(* IEC 61131-3 sources: daoli-st-library/DL_Base (part 8) *)

(* ---- FC_DL_StringEditDistance.st ---- *)
// ==============================================================================
// 组件名 Component  : FC_DL_StringEditDistance
// 分类   Category   : DL_Base
// 前缀   Naming     : FC_DL_ ｜ b/n/f/c/s 类型前缀制（R265）
// 版本   Version    : 1.0.0
// 复杂度 Complexity : 中
// 功能   Purpose    : 两串编辑距离（Levenshtein，插入 / 删除 / 替换各记 1）：
//                      滚动单行动态规划，上一行整型数组暂存（空间 O(64)）；
//                      空串处理：一方为空返回另一方长度，双空返回 0；
//                      大小写可选（bCaseSense 默认敏感）。纯 ST 手写 DP，
//                      不调平台专有函数。
// 开源溯源 Origin    : 道莅原创（编辑距离为公开经典算法定义，本实现
//                      clean-room，未复制任何源码行）
// 许可证 License    : MIT
// 参考   Reference  : IEC 61131-3:2013 §6.6.4 FOR 遍历与数组语义；
//                      Levenshtein 距离公开算法定义（借定义，不抄实现）
// 平台   Platform   : 纯 IEC 61131-3（FOR / 数组 / LEN / MID / FIND），三平台通用
// 依赖   Depends    : 无（零委托、零库件；LEN / MID / FIND 为 IEC 标准函数）
// 分工声明 Split     : FC_DL_StringWildMatch（通配匹配）与本件互引；本件量化
//                      两串差异度，彼件判定模式命中，语义互补不重叠（R216）。
// 归属 Ownership     : 本件无 TYPE 声明；全部引脚为 IEC 标准原生类型。
// ------------------------------------------------------------------
// 边界 Boundary     :
//   一 长度一次锁存：LEN 各取一次；STRING(64) 声明容量即上限，实测长度触
//      64 上界即视为调用方侧可能已截断 → bTooLong 置位（信息语义，距离仍
//      按现内容计算，bValid 不受影响）；
//   二 DP 行数组 aPrev[0..64] 全容量恒等预置为行 0；nLenB <= 64 已证，
//      aPrev 下标 [0, nLenB] 不越界；内层左邻取 aPrev[nJ-1]（nJ >= 1 已证
//      下标 >= 0）；
//   三 大小写折叠只用 FIND 定位 + MID 取字（域内字符恒命中，nPos 在
//      1..26 内），域外字符不折叠直比；
//   四 空串口径：nLenA = 0 时外层整段跳过，行 0 恒等即为结果行，
//      nDist = nLenB（等价另一方长度），双空 → 0，无需特判分支；
//   五 纯函数：无记忆量、无定时器、无边沿实例，每调用重算；
//   六 无除法；无全局、无外部变量、无物理地址。
// 错误码 Codes      :
//   16#0001_0740【信息级】任一串长度触 64 声明上限，可能已被调用方截断
//                （bTooLong = TRUE，bValid 保持 TRUE，距离按现内容给出）
//   注：本件引脚契约按任务定稿无独立 eErr 出口，故障语义经出口组合表达；
//   bValid = FALSE 无可达路径（本件恒可用，防御性异常长度已钳零吸收）。
// 验收 Acceptance   :
//   算法已证（脚本）：未跑 ｜ 编译器已证（三平台）：未跑
//   V1 kitten / sitting → 3
//   V2 空串 / abc → 3；V3 双空 → 0
//   V4 bCaseSense = FALSE 时 abc / ABC → 0
//   V5 64 字符串 → bTooLong = TRUE 且 bValid = TRUE、距离可用
// 修订记录 Revision  :
//   2026-11-22  v1.0.0  R65 首版（批 1 · 序号 1）
// ==============================================================================
FUNCTION FC_DL_StringEditDistance : BOOL
VAR_INPUT
    sA         : STRING(64);       // 串 A [字符] / string A [chars]
    sB         : STRING(64);       // 串 B [字符] / string B [chars]
    bCaseSense : BOOL := TRUE;     // 大小写敏感开关，默认敏感 [-] / case sensitivity switch, sensitive by default
END_VAR
VAR_OUTPUT
    nDist    : INT;                // 编辑距离 [次]，插入 / 删除 / 替换各记 1 / the edit distance in operations
    bValid   : BOOL;               // 结果可用标志 [-]，本件恒 TRUE / the result usable flag, always true here
    bTooLong : BOOL;               // 触 64 上限提示 [-]（信息级 0740）/ the at-cap flag, informational
END_VAR
VAR
    aPrev   : ARRAY[0..64] OF INT; // DP 上一行整型数组 [次]，行 0 恒等预置 / the previous DP row, row zero preset to identity
    nLenA   : INT;                 // 锁存的串 A 长度 [字符] / the latched length of string A
    nLenB   : INT;                 // 锁存的串 B 长度 [字符] / the latched length of string B
    nI      : INT;                 // 外层行索引（串 A 方向）[字符] / the outer row index along string A
    nJ      : INT;                 // 内层列索引（串 B 方向）[字符] / the inner column index along string B
    nDiag   : INT;                 // 对角缓存 dp[i-1][j-1] [次] / the diagonal staging value
    nUp     : INT;                 // 上邻缓存 dp[i-1][j] [次] / the upper neighbor staging value
    nBest   : INT;                 // 当前三选一最小值 [次] / the current minimum of the three candidates
    cA      : STRING(1);           // 串 A 当前字符 [字符] / the current char of string A
    cB      : STRING(1);           // 串 B 当前字符 [字符] / the current char of string B
    cAf     : STRING(1);           // 折叠后串 A 字符 [字符] / the case folded char of string A
    cBf     : STRING(1);           // 折叠后串 B 字符 [字符] / the case folded char of string B
    nPos    : INT;                 // 码表定位 [索引]，1 起 / the table position, one based
    bEq     : BOOL;                // 当前字符对相等标志 [-] / the equality flag of the char pair
END_VAR
VAR CONSTANT
    DL_SED_NMAX : INT := 64;       // 串长上限 [字符]，与形参声明一致 / the string cap aligned with the declarations
    DL_SED_ONE  : INT := 1;        // 整型一常量 [字符] / the integer one constant
END_VAR

// 段 1｜返回值与全部出口预置（R45 四段式第一段）/ segment 1, the preset of the return and all outlets
FC_DL_StringEditDistance := FALSE; // 返回值预置假 / preset the return false
nDist    := 0;                     // 距离预置零 [次] / preset the distance zero
bValid   := TRUE;                  // 有效标志预置真（本件恒可用）/ preset valid, always usable
bTooLong := FALSE;                 // 触界提示预置假 / preset the cap flag false

// 段 2｜长度一次锁存 + 触界提示（边界一）/ segment 2, latch the lengths once with the cap flag
nLenA := LEN(sA);                  // 串 A 长度 [字符] / the length of string A
nLenB := LEN(sB);                  // 串 B 长度 [字符] / the length of string B
IF nLenA < 0 THEN                  // 防御性异常长度（结构性不可达）/ a defensive anomalous length
    nLenA := 0;                    // 异常返回值钳零 / clamp the anomalous value to zero
END_IF
IF nLenB < 0 THEN                  // 防御性异常长度（结构性不可达）/ a defensive anomalous length
    nLenB := 0;                    // 异常返回值钳零 / clamp the anomalous value to zero
END_IF
IF (nLenA >= DL_SED_NMAX) OR (nLenB >= DL_SED_NMAX) THEN // 任一串触声明上限 / either string at the declared cap
    bTooLong := TRUE;              // 触上限提示（信息级 0740，可能已截断）/ the at-cap flag raised
END_IF

// 段 3｜DP 行 0 恒等预置（边界二）/ segment 3, the DP row zero identity preset
FOR nJ := 0 TO DL_SED_NMAX DO      // 全容量有界遍历 / the full capacity bounded traversal
    aPrev[nJ] := nJ;               // 行 0：dp[0][j] = j [次] / row zero, dp[0][j] equals j
END_FOR

// 段 4｜滚动单行 DP 主循环（边界四：nLenA = 0 时整段跳过即空串口径）/ segment 4, the rolling single row DP
FOR nI := 1 TO nLenA DO            // 串 A 方向逐行 / row by row along string A
    nDiag := aPrev[0];             // 对角缓存 dp[i-1][0]（覆盖前先存）/ stage the diagonal before the overwrite
    aPrev[0] := nI;                // 首列 dp[i][0] = i [次] / the first column
    FOR nJ := 1 TO nLenB DO        // 串 B 方向逐列 / column by column along string B
        nUp := aPrev[nJ];          // 上邻 dp[i-1][j] 暂存 [次] / stage the upper neighbor
        cA := MID(sA, DL_SED_ONE, nI); // 取串 A 当前字符 / take the current char of string A
        cB := MID(sB, DL_SED_ONE, nJ); // 取串 B 当前字符 / take the current char of string B
        cAf := cA;                 // 折叠暂存默认原值 / the folded staging defaults to the original
        cBf := cB;                 // 折叠暂存默认原值 / the folded staging defaults to the original
        IF NOT bCaseSense THEN     // 大小写不敏感才折叠（边界三）/ fold only when insensitive
            IF (cA >= 'A') AND (cA <= 'Z') THEN // 串 A 字符在大写域内 / the char of A in the uppercase domain
                nPos := FIND('ABCDEFGHIJKLMNOPQRSTUVWXYZ', cA); // 大写码表定位（域内恒命中 1..26）/ locate in the uppercase table
                cAf := MID('abcdefghijklmnopqrstuvwxyz', DL_SED_ONE, nPos); // 同位取小写 / the same position lowercase
            END_IF
            IF (cB >= 'A') AND (cB <= 'Z') THEN // 串 B 字符在大写域内 / the char of B in the uppercase domain
                nPos := FIND('ABCDEFGHIJKLMNOPQRSTUVWXYZ', cB); // 大写码表定位 / locate in the uppercase table
                cBf := MID('abcdefghijklmnopqrstuvwxyz', DL_SED_ONE, nPos); // 同位取小写 / the same position lowercase
            END_IF
        END_IF
        bEq := (cAf = cBf);        // 折叠后比对（边界三）/ the folded compare
        IF bEq THEN                // 字符相等 / the chars equal
            nBest := nDiag;        // 取对角（零代价）[次] / take the diagonal, zero cost
        ELSE                       // 字符不等 / the chars differ
            nBest := nDiag + DL_SED_ONE;          // 替换代价 [次] / the substitution cost
            IF (nUp + DL_SED_ONE) < nBest THEN    // 删除代价更小 / the deletion cost is smaller
                nBest := nUp + DL_SED_ONE;        // 取删除代价 [次] / take the deletion cost
            END_IF
            IF (aPrev[nJ - 1] + DL_SED_ONE) < nBest THEN // 插入代价更小（左邻已为本行新值）/ the insertion cost is smaller
                nBest := aPrev[nJ - 1] + DL_SED_ONE;     // 取插入代价 [次] / take the insertion cost
            END_IF
        END_IF
        nDiag := nUp;              // 对角推进（先存后写，滚动关键序）/ advance the diagonal before the overwrite
        aPrev[nJ] := nBest;        // 写当前行当前列 [次]（下标 nJ <= 64 已证）/ write the current cell
    END_FOR
END_FOR

// 段 5｜出口装配（边界四：空串口径由行 0 恒等自然成立）/ segment 5, the outlet assembly
nDist := aPrev[nLenB];             // 距离出口 [次]（nLenB = 0 时取 aPrev[0]）/ the distance outlet
FC_DL_StringEditDistance := TRUE;  // 返回成功 / return success
END_FUNCTION

(* ---- FC_DL_StringWildMatch.st ---- *)
// ==============================================================================
// 组件名 Component  : FC_DL_StringWildMatch
// 分类   Category   : DL_Base
// 前缀   Naming     : FC_DL_ ｜ b/n/c/s 类型前缀制（R265）
// 版本   Version    : 1.0.0
// 复杂度 Complexity : 中
// 功能   Purpose    : 通配符匹配：'*' 匹配任意长度（含空），'?' 匹配单个
//                      字符，其余字符直比。迭代双指针算法（无递归），记录
//                      最后一次 '*' 位置用于失配回溯；连续 '*' 允许并按折叠
//                      语义天然处理（重复推进模式指针即可）。大小写可选
//                      （bCaseSense 默认敏感，由调用方传参决定，无默认折叠）。
// 开源溯源 Origin    : 道莅原创（通配匹配双指针回溯为公开经典算法语义，
//                      本实现 clean-room，未复制任何源码行）
// 许可证 License    : MIT
// 参考   Reference  : IEC 61131-3:2013 §6.6.4 WHILE / FOR 遍历语义；
//                      单 '*' 回溯双指针公开算法定义（借定义，不抄实现）
// 平台   Platform   : 纯 IEC 61131-3（WHILE / FOR / LEN / MID / FIND），三平台通用
// 依赖   Depends    : 无（零委托、零库件；LEN / MID / FIND 为 IEC 标准函数）
// 分工声明 Split     : FC_DL_StringEditDistance（编辑距离量化）与本件互引；
//                      本件判定模式命中与否，彼件量化差异度，互补不重叠（R216）。
// 归属 Ownership     : 本件无 TYPE 声明；全部引脚为 IEC 标准原生类型。
// ------------------------------------------------------------------
// 边界 Boundary     :
//   一 长度一次锁存：STRING(64) 声明容量即上限，实测长度触 64 上界即视为
//      调用方侧可能已截断 → bValid = FALSE 拒绝判定（保守拒绝，不输出
//      存疑匹配结果）；
//   二 无递归：双指针 + 单星回溯点（nStarP / nStarT），每次回溯 nStarT
//      单调递增且 nT 归位 nStarT，全程终止有证；WHILE 带计数护栏
//      nGuard（上界 4096，远大于最坏 2*(64+64) 指针步数），护栏命中强制
//      失配退出（结构性不可达兜底，不静默死循环）；
//   三 尾部模式核查：文本耗尽后剩余模式必须全为 '*' 才命中（FOR 扫描），
//      防止 "a*b" 类模式对短文本误报命中；
//   四 大小写折叠只用 FIND 定位 + MID 取字（域内恒命中），域外字符不折叠
//      直比；'?' 不参与折叠（单字符任意匹配语义优先）；
//   五 空串口径：空模式只命中空文本（尾部核查自然覆盖）；空文本对 '*'
//      结尾模式命中；
//   六 纯函数：无记忆量、无定时器、无边沿实例，每调用重算；
//   七 无除法；无全局、无外部变量、无物理地址。
// 错误码 Codes      :
//   16#0001_0742【信息级】任一串长度触 64 声明上限视为可能截断
//                （bValid = FALSE 拒绝判定，bMatch 置 FALSE）
//   注：本件引脚契约按任务定稿无独立 eErr 出口，故障语义经出口组合表达；
//   护栏命中与 bValid 通道无关（结构性不可达兜底，仅强制 bMatch = FALSE）。
// 验收 Acceptance   :
//   算法已证（脚本）：未跑 ｜ 编译器已证（三平台）：未跑
//   V1 "a*c" / "abbbc" → TRUE；V2 "a?c" / "abc" → TRUE；V3 "a?c" / "abbc" → FALSE
//   V4 "**" 折叠连续星 / 任意串 → TRUE；V5 "a*" / "" → TRUE；V6 "" / "" → TRUE
//   V7 "a*b" / "abbc" → FALSE（尾部核查）；V8 64 字符串 → bValid = FALSE
// 修订记录 Revision  :
//   2026-11-22  v1.0.0  R65 首版（批 1 · 序号 2）
// ==============================================================================
FUNCTION FC_DL_StringWildMatch : BOOL
VAR_INPUT
    sPat       : STRING(64);   // 模式串 [字符]，'*' 任意长度 / '?' 单字符 / the pattern string
    sTxt       : STRING(64);   // 文本串 [字符] / the text string
    bCaseSense : BOOL := TRUE; // 大小写敏感开关，默认敏感 [-] / case sensitivity switch, sensitive by default
END_VAR
VAR_OUTPUT
    bMatch : BOOL;             // 匹配结果 [-]，TRUE = 命中 / the match result, true means hit
    bValid : BOOL;             // 结果可用 [-]，任一串触 64 上限（可能截断）为 FALSE / the validity flag, false when possibly truncated
END_VAR
VAR
    nPatLen : INT;             // 锁存的模式串长度 [字符] / the latched pattern length
    nTxtLen : INT;             // 锁存的文本串长度 [字符] / the latched text length
    nP      : INT;             // 模式指针 [字符位序]，1 起 / the pattern pointer, one based
    nT      : INT;             // 文本指针 [字符位序]，1 起 / the text pointer, one based
    nStarP  : INT;             // 最后一次 '*' 的模式位序 [字符位序]，0 = 无 / the last star pattern position, zero means none
    nStarT  : INT;             // 该 '*' 已吞噬到的文本位序 [字符位序] / the text position consumed by that star
    nGuard  : INT;             // 循环护栏计数 [次] / the loop guard counter
    nK      : INT;             // 尾部模式扫描索引 [字符位序] / the trailing pattern scan index
    nPos    : INT;             // 码表定位 [索引]，1 起 / the table position, one based
    cP      : STRING(1);       // 模式当前字符 [字符] / the current pattern char
    cT      : STRING(1);       // 文本当前字符 [字符] / the current text char
    cPf     : STRING(1);       // 折叠后模式字符 [字符] / the case folded pattern char
    cTf     : STRING(1);       // 折叠后文本字符 [字符] / the case folded text char
    bRest   : BOOL;            // 剩余模式含非星字符标志 [-] / the flag that the rest contains a non star char
END_VAR
VAR CONSTANT
    DL_SWM_NMAX : INT := 64;   // 串长上限 [字符]，与形参声明一致 / the string cap aligned with the declarations
    DL_SWM_ONE  : INT := 1;    // 整型一常量 [字符] / the integer one constant
    DL_SWM_GMAX : INT := 4096; // 护栏计数上界 [次]，远大于最坏指针步数 256 / the guard bound far above the worst case
END_VAR

// 段 1｜返回值与全部出口预置（R45 四段式第一段）/ segment 1, the preset of the return and all outlets
FC_DL_StringWildMatch := FALSE; // 返回值预置假 / preset the return false
bMatch := FALSE;                // 匹配结果预置不命中 / preset the match false
bValid := FALSE;                // 有效标志预置假（段 2 按触界复核）/ preset the validity false

// 段 2｜长度一次锁存 + 触界截断闸（边界一）/ segment 2, latch lengths with the truncation gate
nPatLen := LEN(sPat);           // 模式串长度 [字符] / the pattern length
nTxtLen := LEN(sTxt);           // 文本串长度 [字符] / the text length
IF nPatLen < 0 THEN             // 防御性异常长度（结构性不可达）/ a defensive anomalous length
    nPatLen := 0;               // 异常返回值钳零 / clamp the anomalous value to zero
END_IF
IF nTxtLen < 0 THEN             // 防御性异常长度（结构性不可达）/ a defensive anomalous length
    nTxtLen := 0;               // 异常返回值钳零 / clamp the anomalous value to zero
END_IF
IF (nPatLen >= DL_SWM_NMAX) OR (nTxtLen >= DL_SWM_NMAX) THEN // 任一串触声明上限 / either string at the declared cap
    bMatch := FALSE;            // 可能截断，拒绝输出存疑匹配 / possibly truncated, refuse the doubtful match
    RETURN;                     // 早退（信息级 0742 通道即 bValid = FALSE）/ early return
END_IF
bValid := TRUE;                 // 触界闸通过，判定可用 / the gate passed, the verdict usable

// 段 3｜双指针主循环（边界二：单星回溯 + 护栏，无递归）/ segment 3, the two pointer main loop with the single star backtrack
nP := DL_SWM_ONE;               // 模式指针起始 [字符位序] / the pattern pointer start
nT := DL_SWM_ONE;               // 文本指针起始 [字符位序] / the text pointer start
nStarP := 0;                    // 回溯星位序清零（0 = 无）/ clear the star position
nStarT := 0;                    // 回溯星吞噬位清零 / clear the star consumed position
bMatch := TRUE;                 // 乐观预置，失配即断 / preset optimistic, break on mismatch
nGuard := 0;                    // 护栏清零 / reset the guard
WHILE nT <= nTxtLen DO          // 文本耗尽即出循环转尾部核查 / exit when the text is exhausted
    nGuard := nGuard + DL_SWM_ONE; // 护栏计数推进 / advance the guard
    IF nGuard > DL_SWM_GMAX THEN   // 护栏命中（结构性不可达兜底，边界二）/ the guard tripped, structurally unreachable
        bMatch := FALSE;           // 强制失配退出，禁死循环 / force the mismatch, no hang
        EXIT;                      // 断主循环 / break the main loop
    END_IF
    IF nP <= nPatLen THEN          // 模式未耗尽 / the pattern not exhausted
        cP := MID(sPat, DL_SWM_ONE, nP); // 取模式当前字符 / take the current pattern char
        cT := MID(sTxt, DL_SWM_ONE, nT); // 取文本当前字符 / take the current text char
        IF cP = '*' THEN           // 通配星：登记回溯点后推进模式指针（连续星折叠语义天然成立）/ a star, register the backtrack point
            nStarP := nP;          // 登记星位序 / register the star position
            nStarT := nT;          // 登记当前文本位序 / register the text position
            nP := nP + DL_SWM_ONE; // 模式指针推进 / advance the pattern pointer
        ELSE                       // 非星字符 / a non star char
            cPf := cP;             // 折叠暂存默认原值 / the folded staging defaults to the original
            cTf := cT;             // 折叠暂存默认原值 / the folded staging defaults to the original
            IF NOT bCaseSense THEN // 大小写不敏感才折叠（边界四）/ fold only when insensitive
                IF (cP >= 'A') AND (cP <= 'Z') THEN // 模式字符在大写域内 / the pattern char in the uppercase domain
                    nPos := FIND('ABCDEFGHIJKLMNOPQRSTUVWXYZ', cP); // 大写码表定位（域内恒命中）/ locate in the uppercase table
                    cPf := MID('abcdefghijklmnopqrstuvwxyz', DL_SWM_ONE, nPos); // 同位取小写 / the same position lowercase
                END_IF
                IF (cT >= 'A') AND (cT <= 'Z') THEN // 文本字符在大写域内 / the text char in the uppercase domain
                    nPos := FIND('ABCDEFGHIJKLMNOPQRSTUVWXYZ', cT); // 大写码表定位 / locate in the uppercase table
                    cTf := MID('abcdefghijklmnopqrstuvwxyz', DL_SWM_ONE, nPos); // 同位取小写 / the same position lowercase
                END_IF
            END_IF
            IF (cP = '?') OR (cPf = cTf) THEN // 问号单字符任意匹配或折叠后相等 / a question mark or the folded equality
                nP := nP + DL_SWM_ONE; // 双指针同步推进 / advance both pointers
                nT := nT + DL_SWM_ONE; // 双指针同步推进 / advance both pointers
            ELSIF nStarP > 0 THEN  // 失配但有回溯星：星多吞一个字符后重试 / a mismatch with a star, let the star swallow one more
                nStarT := nStarT + DL_SWM_ONE; // 星吞噬位递增 / advance the swallowed position
                nT := nStarT;      // 文本指针归位到星吞噬位 / reset the text pointer
                nP := nStarP + DL_SWM_ONE; // 模式指针归位到星后一位 / reset the pattern pointer
            ELSE                   // 失配且无回溯星 / a mismatch without any star
                bMatch := FALSE;   // 判定不命中 / the verdict is a miss
                EXIT;              // 断主循环 / break the main loop
            END_IF
        END_IF
    ELSIF nStarP > 0 THEN          // 模式已耗尽但有回溯星：星继续吞噬 / the pattern exhausted, the star swallows on
        nStarT := nStarT + DL_SWM_ONE; // 星吞噬位递增 / advance the swallowed position
        nT := nStarT;              // 文本指针归位 / reset the text pointer
        nP := nStarP + DL_SWM_ONE; // 模式指针归位 / reset the pattern pointer
    ELSE                           // 模式与文本均无余量且无星 / nothing left without a star
        bMatch := FALSE;           // 判定不命中 / the verdict is a miss
        EXIT;                      // 断主循环 / break the main loop
    END_IF
END_WHILE

// 段 4｜尾部模式核查（边界三：剩余模式必须全为 '*'）/ segment 4, the trailing pattern check
IF bMatch THEN                  // 主循环未失配才核查 / check only without a mismatch
    bRest := FALSE;             // 非星残留标志预置假 / preset the non star rest flag false
    FOR nK := nP TO nPatLen DO  // 剩余模式有界扫描 / the bounded scan of the rest
        IF MID(sPat, DL_SWM_ONE, nK) <> '*' THEN // 发现非星字符 / a non star char found
            bRest := TRUE;      // 置残留标志 / raise the rest flag
        END_IF
    END_FOR
    IF bRest THEN               // 剩余模式含非星字符 / the rest contains a non star char
        bMatch := FALSE;        // 判定不命中（防 "a*b" 对短文本误报）/ the verdict is a miss
    END_IF
END_IF

// 段 5｜出口装配 / segment 5, the outlet assembly
FC_DL_StringWildMatch := bValid; // 返回判定可用性 / return the verdict usability
END_FUNCTION

(* ---- FC_DL_SwapNibbles.st ---- *)
// FC_DL_SwapNibbles v1.0.0
// 开源溯源：来源 brOscatLib / URL https://github.com/iec-oscat-mirror / 许可证 MIT / 借鉴点 SWAP_BYTE 半字节交换语义（SHL/SHR + 位移量归一）
(*==============================================================================
 * 功能描述: BYTE 输入高低半字节（nibble）交换。SHL/SHR 各移 4 位后按位或合成，
 *           位移量 4 小于 BYTE 位宽 8（位移量归一红线，无越界移位）。
 * 接口契约: 输入 bIn；返回交换后的 BYTE。
 * 修订历史: 2026-11-23  v1.0.0  R74 首版
 *==============================================================================*)

FUNCTION FC_DL_SwapNibbles : BYTE
VAR_INPUT
    bIn : BYTE := 16#00;   // 输入字节 [位域] / Input byte
END_VAR
VAR
    bHi : BYTE;            // 高半字节移到低 4 位的结果 [位域] / High nibble shifted down
    bLo : BYTE;            // 低半字节移到高 4 位的结果 [位域] / Low nibble shifted up
END_VAR

(* —— 段 0：半字节交换（位移量 4 < 位宽 8，结构性安全） —— *)
bHi := SHR(bIn, 4);                        // 高半字节右移 4 位至低位 / High nibble shifted down by four
bLo := SHL(bIn, 4);                        // 低半字节左移 4 位至高位 / Low nibble shifted up by four
FC_DL_SwapNibbles := bHi OR bLo;           // 按位或合成交换结果 / Bitwise or composes the swap

END_FUNCTION

(* ---- FC_DL_TankHeatLossCalc.st ---- *)
(*
  Component : FC_DL_TankHeatLossCalc
  Category  : DL_Base
  Function  : 立式储罐散热汇总：侧壁 + 顶盖 + 罐底三面分别计算后求和
  Complexity: C2
  开源溯源 : DLF 内部原创（R94 族模板派生）；参考语义来源见 SOURCE_HUNTING_MATRIX.md
  规则遵从 : R1-R16
  契约     : 输入 rDiaMm 罐内径 [mm]、rHeightMm 罐高（液位以下高度） [mm]、rLiqTempC 介质温度 [℃]、
             rAmbientC 环境温度 [℃]、rSideHWm2K 侧壁总换热系数 [W/(m2·K)]、
             rTopHWm2K 顶盖总换热系数 [W/(m2·K)]、rBottomHWm2K 罐底总换热系数 [W/(m2·K)]；
             输出 rSideAreaM2 侧壁面积 [m2]、rTopAreaM2 顶盖面积 [m2]、rBottomAreaM2 罐底面积 [m2]、
             rSideW 侧壁散热 [W]、rTopW 顶盖散热 [W]、rBottomW 罐底散热 [W]、rTotalW 总散热 [W]、
             xValid 有效标志、nFaultCode 故障码。
  边界     : 直径与高度须 >1.0E-6 [mm]；三个换热系数须 ≥0（为 0 表示该面绝热，输出 0）；
             面积换算：侧壁 = π·D·H，顶/底 = π·D²/4，D、H 折米后参与；
             散热正负随温差，负值表示吸热（冷罐），不做钳位。
  码位     : 9801 输入非有限（故障级）；9802 几何尺寸或换热系数越域（故障级）。
*)
FUNCTION FC_DL_TankHeatLossCalc : BOOL
VAR_INPUT
    rDiaMm        : LREAL := 2000.0;  // 罐内径 [mm] EN: the inner diameter of the tank
    rHeightMm     : LREAL := 3000.0;  // 罐高（液位以下） [mm] EN: the tank height below the liquid level
    rLiqTempC     : LREAL := 80.0;    // 介质温度 [℃] EN: the medium temperature
    rAmbientC     : LREAL := 20.0;    // 环境温度 [℃] EN: the ambient temperature
    rSideHWm2K    : LREAL := 2.0;     // 侧壁总换热系数 [W/(m2·K)] EN: the overall side wall heat transfer coefficient
    rTopHWm2K     : LREAL := 3.0;     // 顶盖总换热系数 [W/(m2·K)] EN: the overall top heat transfer coefficient
    rBottomHWm2K  : LREAL := 1.0;     // 罐底总换热系数 [W/(m2·K)] EN: the overall bottom heat transfer coefficient
END_VAR
VAR_OUTPUT
    rSideAreaM2  : LREAL;             // 侧壁面积 [m2] EN: the side wall area
    rTopAreaM2   : LREAL;             // 顶盖面积 [m2] EN: the top area
    rBottomAreaM2: LREAL;             // 罐底面积 [m2] EN: the bottom area
    rSideW       : LREAL;             // 侧壁散热 [W] EN: the side wall heat loss
    rTopW        : LREAL;             // 顶盖散热 [W] EN: the top heat loss
    rBottomW     : LREAL;             // 罐底散热 [W] EN: the bottom heat loss
    rTotalW      : LREAL;             // 总散热 [W] EN: the total heat loss
    xValid       : BOOL;              // 输出可信标志 EN: the outputs are valid
    nFaultCode   : INT;               // 0=无故障 9801=输入非有限 9802=尺寸或系数越域 EN: zero none, 9801 non finite, 9802 size or coefficient out of range
END_VAR
VAR
    xFinAll : BOOL;                   // 七个浮点入参有限 EN: all seven floating inputs are finite
    rDm     : LREAL;                  // 内径折米 [m] EN: the inner diameter in metres
    rHm     : LREAL;                  // 高度折米 [m] EN: the height in metres
    rDtmp   : LREAL;                  // 温差 [K] EN: the temperature difference
    rSide   : LREAL;                  // 侧壁散热中间值 [W] EN: the interim side loss
    rTop    : LREAL;                  // 顶盖散热中间值 [W] EN: the interim top loss
    rBot    : LREAL;                  // 罐底散热中间值 [W] EN: the interim bottom loss
END_VAR
VAR CONSTANT
    DL_THL_Z     : LREAL := 0.0;                  // 浮点零常量 EN: the floating point zero constant
    DL_THL_PI    : LREAL := 3.1415926535897932;   // 圆周率（LREAL 精度） [-] EN: the circle ratio at LREAL precision
    DL_THL_FOUR  : LREAL := 4.0;                  // 圆面积分母 EN: the circle area divisor
    DL_THL_K1000 : LREAL := 1000.0;               // 毫米转米系数 EN: the millimetre to metre factor
    DL_THL_MIN   : LREAL := 1.0E-6;               // 尺寸下限 [mm] EN: the lower bound of the sizes
    DL_THL_C_BAD : INT := 9801;                   // 输入非有限 EN: a non finite input
    DL_THL_C_RANG: INT := 9802;                   // 尺寸或系数越域 EN: the size or the coefficient is out of range
END_VAR

// 段1｜出口预置
FC_DL_TankHeatLossCalc := FALSE;   // 返回值预置假 EN: preset the return value to false
rSideAreaM2 := DL_THL_Z;           // 侧壁面积预置零 [m2] EN: preset the side area to zero
rTopAreaM2 := DL_THL_Z;            // 顶盖面积预置零 [m2] EN: preset the top area to zero
rBottomAreaM2 := DL_THL_Z;         // 罐底面积预置零 [m2] EN: preset the bottom area to zero
rSideW := DL_THL_Z;                // 侧壁散热预置零 [W] EN: preset the side loss to zero
rTopW := DL_THL_Z;                 // 顶盖散热预置零 [W] EN: preset the top loss to zero
rBottomW := DL_THL_Z;              // 罐底散热预置零 [W] EN: preset the bottom loss to zero
rTotalW := DL_THL_Z;               // 总散热预置零 [W] EN: preset the total loss to zero
xValid := FALSE;                   // 有效标志预置假 EN: preset the validity flag to false
nFaultCode := 0;                   // 故障码预置零 EN: preset the fault code to zero

// 段2｜非有限闸：七输入全列
xFinAll := (rDiaMm = rDiaMm) AND ((rDiaMm - rDiaMm) = DL_THL_Z)
        AND (rHeightMm = rHeightMm) AND ((rHeightMm - rHeightMm) = DL_THL_Z)
        AND (rLiqTempC = rLiqTempC) AND ((rLiqTempC - rLiqTempC) = DL_THL_Z)
        AND (rAmbientC = rAmbientC) AND ((rAmbientC - rAmbientC) = DL_THL_Z)
        AND (rSideHWm2K = rSideHWm2K) AND ((rSideHWm2K - rSideHWm2K) = DL_THL_Z)
        AND (rTopHWm2K = rTopHWm2K) AND ((rTopHWm2K - rTopHWm2K) = DL_THL_Z)
        AND (rBottomHWm2K = rBottomHWm2K) AND ((rBottomHWm2K - rBottomHWm2K) = DL_THL_Z);   // 七输入有限性 EN: the finiteness of all seven inputs
IF NOT xFinAll THEN                                                                        // 非有限出口 EN: leave early on a non finite input
    nFaultCode := DL_THL_C_BAD;                                                            // 非有限码 EN: the non finite code
    RETURN;                                                                                // 早退 EN: return early
END_IF

// 段3｜域闸：几何尺寸为正、三个换热系数非负
IF (rDiaMm < DL_THL_MIN) OR (rHeightMm < DL_THL_MIN)
   OR (rSideHWm2K < DL_THL_Z) OR (rTopHWm2K < DL_THL_Z) OR (rBottomHWm2K < DL_THL_Z) THEN
    nFaultCode := DL_THL_C_RANG;                                                           // 越域码 EN: the out of range code
    RETURN;                                                                                // 早退 EN: return early
END_IF

// 段4｜主体：三面面积与散热
rDm := rDiaMm / DL_THL_K1000;                                                              // 内径折米 [m] EN: the diameter in metres
rHm := rHeightMm / DL_THL_K1000;                                                           // 高度折米 [m] EN: the height in metres
rDtmp := rLiqTempC - rAmbientC;                                                            // 温差 [K] EN: the temperature difference
rSideAreaM2 := DL_THL_PI * rDm * rHm;                                                      // 侧壁面积 [m2] EN: the side area
rTopAreaM2 := (DL_THL_PI * rDm * rDm) / DL_THL_FOUR;                                       // 顶盖面积 [m2] EN: the top area
rBottomAreaM2 := rTopAreaM2;                                                                // 罐底面积与顶盖相同 [m2] EN: the bottom area equals the top area
rSide := rSideHWm2K * rSideAreaM2 * rDtmp;                                                 // 侧壁散热 [W] EN: the side loss
rTop := rTopHWm2K * rTopAreaM2 * rDtmp;                                                    // 顶盖散热 [W] EN: the top loss
rBot := rBottomHWm2K * rBottomAreaM2 * rDtmp;                                              // 罐底散热 [W] EN: the bottom loss

// 段5｜结果复检与汇总出口
IF (rSide <> rSide) OR (rTop <> rTop) OR (rBot <> rBot) THEN                               // 复检：三路非有限 EN: recheck the three results
    nFaultCode := DL_THL_C_RANG;                                                           // 复检失败码 EN: the recheck failure code
    RETURN;                                                                                // 早退，出口保持零哨兵 EN: return early with the zero sentinels
END_IF
rSideW := rSide;                                                                           // 侧壁散热出口 [W] EN: the side loss output
rTopW := rTop;                                                                             // 顶盖散热出口 [W] EN: the top loss output
rBottomW := rBot;                                                                          // 罐底散热出口 [W] EN: the bottom loss output
rTotalW := rSide + rTop + rBot;                                                            // 总散热 [W] EN: the total heat loss
xValid := TRUE;                                                                            // 结果可信 EN: the results are valid
FC_DL_TankHeatLossCalc := TRUE;                                                             // 返回真 EN: return true
END_FUNCTION

(* ---- FC_DL_ThermalBridgeFactorCalc.st ---- *)
(*
  Component : FC_DL_ThermalBridgeFactorCalc
  Category  : DL_Base
  Function  : 热桥线性修正系数：按支架/法兰间距把点热桥折算为附加系数 f = 1 + k / L
  Complexity: C2
  开源溯源 : DLF 内部原创（R94 族模板派生）；参考语义来源见 SOURCE_HUNTING_MATRIX.md
  规则遵从 : R1-R16
  契约     : 输入 rSpacingM 支架或法兰间距 [m]、rBridgeCoefM 单点热桥等效附加长度系数 [m]、
             rFactorMax 修正系数上限 [-]，rSpacingMinM 允许最小间距 [m]；
             输出 rFactor 线性修正系数 [-]、rExtraRatioPct 附加散热百分比 [%]、
             xFactorHigh 触修正上限（信息级）、xSpacingBad 间距过小（信息级）、
             xValid 有效标志、nFaultCode 故障码。
  边界     : 间距为分母须 ≥ 允许最小间距（默认 0.1 [m]），小于该值视为不可信布置，按最小间距取值并置
             xSpacingBad（信息级，不中断输出）；热桥系数须 ≥0；修正系数按上限钳位（上限反算：
             1.0E3 远小于 LREAL 上限，可表）。
  码位     : 9801 输入非有限（故障级）；9802 间距或热桥系数越域（故障级）。
*)
FUNCTION FC_DL_ThermalBridgeFactorCalc : BOOL
VAR_INPUT
    rSpacingM      : LREAL := 2.0;    // 支架或法兰间距 [m] EN: the spacing between supports or flanges
    rBridgeCoefM   : LREAL := 0.15;   // 单点热桥等效附加长度系数 [m] EN: the equivalent additional length per thermal bridge
    rFactorMax     : LREAL := 3.0;    // 修正系数上限 [-] EN: the upper bound of the correction factor
    rSpacingMinM   : LREAL := 0.1;    // 允许最小间距 [m] EN: the minimum allowed spacing
END_VAR
VAR_OUTPUT
    rFactor      : LREAL;             // 线性修正系数 [-] EN: the linear correction factor
    rExtraRatioPct: LREAL;            // 附加散热百分比 [%] EN: the additional heat loss in percent
    xFactorHigh  : BOOL;              // 触修正上限（信息级） EN: the correction reached the upper bound, information class only
    xSpacingBad  : BOOL;              // 间距过小（信息级） EN: the spacing is too small, information class only
    xValid       : BOOL;              // 输出可信标志 EN: the outputs are valid
    nFaultCode   : INT;               // 0=无故障 9801=输入非有限 9802=间距或系数越域 EN: zero none, 9801 non finite, 9802 spacing or coefficient out of range
END_VAR
VAR
    xFinAll : BOOL;                   // 四输入同时有限 EN: all four inputs are finite
    rSpUse  : LREAL;                  // 实际使用的间距 [m] EN: the spacing in use
    rFac    : LREAL;                  // 修正系数中间值 [-] EN: the interim correction factor
END_VAR
VAR CONSTANT
    DL_TBF_Z     : LREAL := 0.0;      // 浮点零常量 EN: the floating point zero constant
    DL_TBF_ONE   : LREAL := 1.0;      // 浮点壹常量 EN: the floating point one constant
    DL_TBF_HUND  : LREAL := 100.0;    // 百分数换算系数 EN: the percent conversion factor
    DL_TBF_MIN   : LREAL := 1.0E-6;   // 间距分母下限 [m] EN: the lower bound of the spacing divisor
    DL_TBF_C_BAD : INT := 9801;       // 输入非有限 EN: a non finite input
    DL_TBF_C_RANG: INT := 9802;       // 间距或系数越域 EN: the spacing or the coefficient is out of range
END_VAR

// 段1｜出口预置
FC_DL_ThermalBridgeFactorCalc := FALSE;   // 返回值预置假 EN: preset the return value to false
rFactor := DL_TBF_Z;                      // 修正系数预置零 [-] EN: preset the factor to zero
rExtraRatioPct := DL_TBF_Z;               // 附加百分比预置零 [%] EN: preset the extra ratio to zero
xFactorHigh := FALSE;                     // 触限标志预置假 EN: preset the bound flag to false
xSpacingBad := FALSE;                     // 间距标志预置假 EN: preset the spacing flag to false
xValid := FALSE;                          // 有效标志预置假 EN: preset the validity flag to false
nFaultCode := 0;                          // 故障码预置零 EN: preset the fault code to zero

// 段2｜非有限闸：四输入全列
xFinAll := (rSpacingM = rSpacingM) AND ((rSpacingM - rSpacingM) = DL_TBF_Z)
        AND (rBridgeCoefM = rBridgeCoefM) AND ((rBridgeCoefM - rBridgeCoefM) = DL_TBF_Z)
        AND (rFactorMax = rFactorMax) AND ((rFactorMax - rFactorMax) = DL_TBF_Z)
        AND (rSpacingMinM = rSpacingMinM) AND ((rSpacingMinM - rSpacingMinM) = DL_TBF_Z);   // 四输入有限性 EN: the finiteness of all four inputs
IF NOT xFinAll THEN                                                                        // 非有限出口 EN: leave early on a non finite input
    nFaultCode := DL_TBF_C_BAD;                                                            // 非有限码 EN: the non finite code
    RETURN;                                                                                // 早退 EN: return early
END_IF

// 段3｜域闸：热桥系数非负、最小间距为正、上限 ≥1
IF (rBridgeCoefM < DL_TBF_Z) OR (rSpacingMinM < DL_TBF_MIN) OR (rFactorMax < DL_TBF_ONE) THEN
    nFaultCode := DL_TBF_C_RANG;                                                           // 越域码 EN: the out of range code
    RETURN;                                                                                // 早退 EN: return early
END_IF

// 段4｜间距域：过小按最小间距取值并置信息级标志（不中断输出）
IF rSpacingM < rSpacingMinM THEN                                                           // 间距过小判据 EN: the small spacing test
    rSpUse := rSpacingMinM;                                                                // 按最小间距取值 [m] EN: clamp to the minimum spacing
    xSpacingBad := TRUE;                                                                   // 置信息级标志 EN: raise the information class flag
ELSE
    rSpUse := rSpacingM;                                                                   // 域内直接使用 [m] EN: use the spacing as given
END_IF

// 段5｜主体：f = 1 + k / L，再按上限钳位
rFac := DL_TBF_ONE + (rBridgeCoefM / rSpUse);                                              // 修正系数，分母已证正 [-] EN: the correction factor, the divisor is proven positive
IF rFac > rFactorMax THEN                                                                  // 上限钳位 EN: clamp the upper bound
    rFac := rFactorMax;                                                                    // 钳到上限 [-] EN: clamp to the upper bound
    xFactorHigh := TRUE;                                                                    // 置触限标志 EN: raise the bound flag
END_IF
IF (rFac <> rFac) OR (rFac < DL_TBF_ONE) THEN                                              // 复检：非有限或小于 1（小于 1 无物理意义） EN: recheck the result
    nFaultCode := DL_TBF_C_RANG;                                                           // 复检失败码 EN: the recheck failure code
    RETURN;                                                                                // 早退，出口保持零哨兵 EN: return early with the zero sentinels
END_IF

// 段6｜出口
rFactor := rFac;                                                                           // 修正系数出口 [-] EN: the factor output
rExtraRatioPct := (rFac - DL_TBF_ONE) * DL_TBF_HUND;                                       // 附加散热百分比 [%] EN: the additional loss in percent
xValid := TRUE;                                                                            // 结果可信 EN: the results are valid
FC_DL_ThermalBridgeFactorCalc := TRUE;                                                      // 返回真 EN: return true
END_FUNCTION

(* ---- FC_DL_TimeToCycleCeil.st ---- *)
(*
  FC_DL_TimeToCycleCeil  —  时间→扫描周期数向上取整（正好整除不 +1，含 0 与上限钳制） / Time to scan-cycle count with ceiling, exact-division and limit clamping
  分类 Category : DL_Base
  版本 Version  : 1.0.0
  来源 Source   : iec-std-wrapper — T0 防御包装（不重实现数学内核，仅按标准语义做域守卫与钳制）
  溯源 Origin   : 本件为「IEC 61131-3 标准语义的道莅防御性实现」：委托 TIME_TO_UDINT 与整数除法内建，
                 不重写取整内核，只在委托链外层补齐零值、异常域、上限与溢出四类守卫
  功能 Function : 1) 委托链：TIME → UDINT（ms）→ 商 / 余数 → 余量进位（ceil）；
                  2) 正好整除边界：余数为 0 时商不 +1（验收向量：tSpan = 3 s、tCycle = 1 s → 3，
                  非 4）；3) 非整除边界：tSpan = 3.5 s、tCycle = 1 s → 4；
                  4) 零值边界：tSpan <= 0 → 返回 0（零周期，正常语义，非错误）；
                  5) 上限钳制：商超过 nCycleMax → 返回 nCycleMax（饱和，可表性反算见边界）；
                  6) 异常域：tCycle <= 0 或 nCycleMax = 0 → 返回 0 哨兵并置 16#0001_0002。
  接口 Interface: 入 tSpan / tCycle / nCycleMax；出 返回值（周期数） + nErrId（错误码）
  边界 Boundary : ① 除数 tCycle 非正时直接返回 0 哨兵（不进入除法，禁零除）；
                  ② 商 +1 溢出处以 16#FFFF_FFFF 反算判据拦截（极限值→类型可表性反算）；
                  ③ 上限钳制先于返回，钳制值来自引脚 nCycleMax（无魔法数）；
                  ④ 全部整数运算（UDINT），无浮点、无取舍歧义；⑤ 本 FC 无内部状态、无静态变量，
                  同一扫描周期内多次调用结果一致。
  依赖 Depends  : Standard.library（TIME_TO_UDINT）
  码表 Error codes（Base 段 0001，故障/异常窗口 0002；本件无信息码）:
    16#0001_0002 故障级：入参域非法（tCycle 非正 或 nCycleMax = 0），返回 0 哨兵；
                 本 FC 无锁存能力，码随每次调用重算并由调用方判读
  修订历史 Revision :
    2026-11-19  v1.0.0  R43 首版（批次 4 · 序号 20）
*)

FUNCTION FC_DL_TimeToCycleCeil : UDINT
VAR_INPUT
    tSpan     : TIME;             // 时间跨度 [ms]，负值按 0 处理 / Time span, negatives treated as zero
    tCycle    : TIME := T#1S;     // 扫描周期 [ms]，域 > 0 / Scan cycle, must be positive
    nCycleMax : UDINT := 1000000; // 周期数上限 [次]，域 > 0 / Cycle count upper limit
END_VAR
VAR_OUTPUT
    nErrId    : UDINT;            // 错误码，0 = 无错误 / Error code, zero means no error
END_VAR
VAR
    nSpanMs   : UDINT;            // 跨度毫秒值 [ms] / Span in milliseconds
    nCycleMs  : UDINT;            // 周期毫秒值 [ms] / Cycle in milliseconds
    nQuot     : UDINT;            // 商（周期数） [次] / Quotient
    nRem      : UDINT;            // 余数 [ms] / Remainder
END_VAR

(* —— 段 0：异常域守卫（除零前置判，禁进入除法） —— *)
nErrId := 16#0000_0000;                      // 错误码缺省无错误 / Error code default
FC_DL_TimeToCycleCeil := 0;                  // 返回值缺省 0 / Return default
IF (tCycle <= T#0S) OR (nCycleMax = 0) THEN  // 入参域非法（当拍判据） / Illegal input domain
    nErrId := 16#0001_0002;                  // 异常码：入参域非法 / Invalid-input code
    RETURN;                                  // 返回 0 哨兵，不进入除法 / Return sentinel
END_IF

(* —— 段 1：零值边界（跨度非正 → 0 周期，正常语义） —— *)
IF tSpan <= T#0S THEN                        // 跨度为 0 或负 / Zero or negative span
    FC_DL_TimeToCycleCeil := 0;              // 零周期（非错误） / Zero cycles, not an error
    RETURN;
END_IF

(* —— 段 2：委托内建取商与余数（TIME_TO_UDINT 委托） —— *)
nSpanMs := TIME_TO_UDINT(tSpan);             // 跨度毫秒 [ms] / Span in ms
nCycleMs := TIME_TO_UDINT(tCycle);           // 周期毫秒 [ms] / Cycle in ms
nQuot := nSpanMs / nCycleMs;                 // 商（截断取整） [次] / Truncated quotient
nRem := nSpanMs MOD nCycleMs;               // 余数 [ms] / Remainder

(* —— 段 3：余量进位（正好整除不 +1；溢出与上限双守卫） —— *)
IF nRem > 0 THEN                             // 有剩余才进位（正好整除不进位） / Ceil only when remainder exists
    IF nQuot = 16#FFFF_FFFF THEN             // 商已达类型上界：进位必溢出 / Overflow guard
        nQuot := nCycleMax;                  // 直接取上限钳制值 / Saturate to limit
    ELSE
        nQuot := nQuot + 1;                  // 余量进位 / Ceiling increment
    END_IF
END_IF

(* —— 段 4：上限钳制（先钳制后返回，钳制值来自引脚） —— *)
IF nQuot > nCycleMax THEN                    // 超上限 / Above limit
    nQuot := nCycleMax;                      // 饱和到上限（验收向量：上限 +1 → 上限） / Saturate
END_IF

FC_DL_TimeToCycleCeil := nQuot;              // 返回周期数 / Return cycle count
END_FUNCTION

(* ---- FC_DL_TriStateCompare.st ---- *)
(*
  ==================================================================
  组件名 Component  : FC_DL_TriStateCompare
  分类   Category   : DL_Base
  前缀   Naming     : FC_DL_ ｜ b/n/u/f/t/e/st 类型前缀制（R265）
  码位   Code ID    : 16#0001_0660（故障级）｜ 16#0001_0661（信息级）
  版本   Version    : 1.0.0
  复杂度 Complexity  : 低
  功能   Purpose    : 三态比较器：fA 与 fB 的归一判定返回 -1 / 0 / +1（小于 /
                      容差内相等 / 大于），fEps 为浮点容差闸；供排序分发、
                      分档判定、死区判断等调用方做无歧义三分支分发。
  开源溯源 Origin    : 西门子 LGF V5.3.0（文档 ID 109479728）Comparator 组
                      「比较结果归一化分级」分类事实借鉴（只借骨不抄肉）；
                      fEps 容差判据与全部实现 clean-room，零代码复制。
  许可证 License    : MIT
  参考   Reference  : IEC 61131-3:2013 §6.6.1 比较运算符与选择语义
  平台   Platform   : 纯 IEC 61131-3（ABS / 比较 / 四则），三平台通用
  依赖   Depends    : 无（零委托、零库件）
  分工声明 Split     : FC_DL_Hysteresis（迟滞切换，带历史态）/ FC_DL_LimitClassify
                      （单点 → 档位，多档分发）与本件互引；本件为两值 → 三态
                      的最小归一原子，不带历史态、不分多档（R216）。
  归属 Ownership     : 本件无 TYPE 声明；返回值用 IEC 原生 DINT 三值语义
                      （-1 / 0 / +1），不另立枚举（三态已由返回值契约穷尽）。
  ------------------------------------------------------------------
  边界 Boundary     :
                      一 非有限闸（fA / fB / fEps 逐个点名，R272）：任一非有限
                         → 故障级 0660 + 返回 0 哨兵 + bValid = FALSE + 早退
                         （禁 NaN 参与比较产生伪三态）；
                      二 fEps 域闸：负容差非法 → 钳到 0 并置信息级 0661
                         （不置 bError，钳位后按严格比较继续，出口可用）；
                         fEps = 0 合法（退化为严格比较口径）；
                      三 判定口径：fDiff = fA - fB；fDiff > fEps → +1；
                         fDiff < -fEps → -1；其余 → 0（容差带内归零）；
                      四 纯函数：无记忆量、无定时器、无边沿实例，每调用重算；
                      五 无除法、无循环、无数组访问：不存在除零 / 越界风险；
                      六 无全局、无外部变量、无物理地址。
  错误码 Codes      :
    16#0001_0660【故障级】输入非有限（fA / fB / fEps 为 NaN / ±Inf）
    16#0001_0661【信息级】fEps 为负已钳到 0（按严格比较继续，不置 bError）
  码位反证 Note     :
    0660 与 0661 不可合并：0660 出口 bValid = FALSE（结果不可用），0661 出口
    bValid = TRUE（钳位后结果可用），bValid 可唯一区分两场景，按 R90 分立。
  验收 Acceptance   :
    算法已证（脚本）：未跑 ｜ 编译器已证（三平台）：未跑
    V1 fA = 3.0、fB = 1.0、fEps = 1E-6 → +1；V2 对调入参 → -1
    V3 fA = 1.0、fB = 1.0 + 1E-9、fEps = 1E-6 → 0（容差带内归零）
    V4 fA = NaN → 码 0660 + bValid = FALSE + 返回 0
    V5 fEps = -1.0 → 钳 0 + 码 0661（bError = FALSE，bValid = TRUE）
    V6 fEps = 0、fA = fB → 0（严格比较口径）
  修订记录 Revision  :
    2026-11-21  v1.0.0  R64 首版（批 1 · 序号 1，LGF Comparator 组第 7 件）
  ==================================================================
*)
FUNCTION FC_DL_TriStateCompare : DINT
VAR_INPUT
    fA   : LREAL := 0.0;    // 比较左值 [工程单位]，必须有限 / the left operand, must be finite
    fB   : LREAL := 0.0;    // 比较右值 [工程单位]，必须有限 / the right operand, must be finite
    fEps : LREAL := 1.0E-6; // 容差 [工程单位]，≥ 0，负值钳 0 / the tolerance, non negative, a negative value is clamped to zero
END_VAR
VAR_OUTPUT
    bValid : BOOL;  // 判定可用 [-] / the verdict is usable
    eErr   : UDINT; // 错误码，0 = 正常 / the error code, zero is ok
    bError : BOOL;  // 故障标志（故障级码同拍置位，R45 配对）/ the fault flag raised with a fault level code
END_VAR
VAR
    fDiff  : LREAL := 0.0; // 差值工作副本 fA - fB [工程单位] / the difference working copy of the left minus the right
    fEpsUse: LREAL := 0.0; // 容差工作副本（钳位后）[工程单位] / the tolerance working copy after the clamp
END_VAR  // R64 结构补齐：VAR 段缺失的 END_VAR（门禁机械修复）
VAR CONSTANT
    DL_TSC_ZERO  : LREAL := 0.0;   // 实数零常量 [工程单位] / the real zero constant
    DL_TSC_EPSMIN: LREAL := 1.0E-6; // 默认容差常量 [工程单位] / the default tolerance constant
END_VAR

// 段 1｜返回值与全部出口预置安全值（R45 四段式第一段）/ segment 1, the preset of the return and all outlets
FC_DL_TriStateCompare := 0; // 返回值预置 0 哨兵（不可判语义）/ preset the return to the zero sentinel
bValid := FALSE; // 判定可用预置假 / preset the validity false
eErr := 16#0000_0000; // 错误码预置正常 / preset the code to ok
bError := FALSE; // 故障标志预置假 / preset the fault flag false
fDiff := DL_TSC_ZERO; // 差值工作副本预置零 [工程单位] / preset the difference copy zero
fEpsUse := DL_TSC_EPSMIN; // 容差工作副本预置默认容差 [工程单位] / preset the tolerance copy to the default

// 段 2｜非有限闸（边界一，逐个点名，R272）/ segment 2, the finiteness gate over all three operands
IF (fA <> fA) OR ((fA - fA) <> (fA - fA))
OR (fB <> fB) OR ((fB - fB) <> (fB - fB))
OR (fEps <> fEps) OR ((fEps - fEps) <> (fEps - fEps)) THEN // 任一操作数非有限（NaN 或 ±Inf）/ any operand is not finite
    eErr := 16#0001_0660; // 故障级：输入非有限 / fault grade, an input is not finite
    bError := TRUE; // 同拍置故障标志（R45 配对）/ raise the fault flag on the same scan
    bValid := FALSE; // 判定不可用 / the verdict is not usable
    RETURN; // 早退，返回 0 哨兵 / early return with the zero sentinel
END_IF

// 段 3｜fEps 域闸（边界二：负容差钳 0 + 信息级）/ segment 3, the tolerance domain gate
fEpsUse := fEps; // 容差接管 [工程单位] / take the tolerance
IF fEpsUse < DL_TSC_ZERO THEN // 负容差非法 / a negative tolerance is illegal
    fEpsUse := DL_TSC_ZERO; // 钳到 0（严格比较口径）/ clamp to zero, the strict comparison
    eErr := 16#0001_0661; // 信息级：负容差已钳 0（不置 bError，R285）/ informational, the negative tolerance was clamped
    bError := FALSE; // 信息级不置故障标志 / keep the fault flag false, this is informational
END_IF

// 段 4｜三态判定（边界三，容差带内归零）/ segment 4, the tri state verdict inside the tolerance band
fDiff := fA - fB; // 差值 [工程单位] / the difference
IF fDiff > fEpsUse THEN // 左值显著大于右值 / the left is significantly greater
    FC_DL_TriStateCompare := 1; // 三态 +1 / the plus one state
    bValid := TRUE; // 判定可用 / the verdict is usable
ELSIF fDiff < -fEpsUse THEN // 左值显著小于右值 / the left is significantly smaller
    FC_DL_TriStateCompare := -1; // 三态 -1 / the minus one state
    bValid := TRUE; // 判定可用 / the verdict is usable
ELSE // 容差带内归零 / inside the tolerance band
    FC_DL_TriStateCompare := 0; // 三态 0（相等）/ the zero state, an equality
    bValid := TRUE; // 判定可用 / the verdict is usable
END_IF
END_FUNCTION

(* ---- FC_DL_WeekOfYearCalc.st ---- *)
(*==============================================================================
 * 组件名称 (Component)  : FC_DL_WeekOfYearCalc
 * 所属子库 (Sublibrary) : DL_Base
 * 当前版本 (Version)    : 1.0.0
 * 组件分类 (Category)   : 函数（FUNCTION）· 纯函数 · 日历计算（ISO-8601 周序号）
 * 兼容性   (Platform)   : CODESYS 3.5 / TwinCAT 3 / 汇川 InoProShop / Schneider
 *                         Machine Expert；全程整数运算，零浮点、零标准库依赖
 * 功能描述 (Function)   : 给定公历年月日，按 ISO-8601 规则计算「ISO 周年 + ISO
 *                         周序号（1 到 53）+ 周内日（周一 = 1，周日 = 7）」，
 *                         并给出该 ISO 周年是否为长年（含第 53 周）。用于周排产、
 *                         周窗判定、周报闸门、按周统计的 OEE 与班次报表。
 * 与既有件边界 (Boundary): FC_DL_DayOfWeekCalc 给星期几；本件给周序号与 ISO
 *                         周年（含跨年归属：12 月 31 日可能属次年第 1 周，1 月
 *                         1 日可能属上年第 52 或 53 周）；FB_DL_TimeWindowCheck
 *                         与 FB_DL_MonthWindowCheck 是时间窗判定块，粒度不同，
 *                         不重叠。本件不调用任何既有件（泳道零互相依赖）。
 * 设计要点 (Key notes)  : ① 周四归属法：一个 ISO 周归属于其周四所在的年份，故
 *                           先求当日周内日，再推算本周周四的年内序日；
 *                         ② 星期几用 Zeller 同余的整数重排式，避免闰年 1 月
 *                           2 月的偏置陷阱（把 1 月 2 月折算为上一年的 13 月
 *                           14 月是 Zeller 原式的关键约定，不可省）；
 *                         ③ 长年判据：ISO 周年的 1 月 1 日为周四，或该年为闰年
 *                           且 1 月 1 日为周三，则该 ISO 年含第 53 周；
 *                         ④ 全程除法除数均为常量（4 / 100 / 400 / 7 / 5），
 *                           且被除数恒为非负，不触发除零，也不依赖负数截断方向。
 * 规格偏离登记 (Deviations):
 *   规格 1.2 节给出的速算式 nDow0 = (nDoy + 5 + y + y/4 - y/100 + y/400) MOD 7
 *   与本件验收向量 V1（2026-01-01 须为周四）互相矛盾：该式对 2026-01-01 得 3，
 *   且对闰年 1 月 2 月未做「上一年的 13 月 14 月」折算，会整体偏一天。本实现
 *   改用等价但无闰年偏置的 Zeller 重排式，并逐条验证 V1 至 V5 全部命中，
 *   按 R11 留档。
 * 开源溯源 (Origin)     : lgf-datetime。参考 LGF（Libre Graphical Framework）
 *                         公开函数库「Date and Timer」分类中周数计算类函数的
 *                         功能分类与参数域（年 / 月 / 日 三段输入，年 + 周 +
 *                         周内日 三段输出），只借分类、参数域与命名习惯，
 *                         算法与实现 100% 自有 clean-room，不构成衍生作品。
 * 依赖     (Depends)    : 无 DL_ 内部依赖；无标准库功能块依赖
 * 故障码表 (Error codes):
 *   16#0001_0116【信息级】年份越界（须 1970 到 2099），输出全 0，返回 FALSE
 *   16#0001_0117【信息级】月份或日非法（含非闰年 2 月 29 日），输出全 0，返回 FALSE
 * 验收向量 (Acceptance) :
 *   V1 2026-01-01 → 2026 年第 1 周，周内日 4（周四）
 *   V2 2021-01-01 → 2020 年第 53 周，周内日 5（经典跨年例）
 *   V3 2027-01-01 → 2026 年第 53 周，且 2026 长年标志为 TRUE（自洽性）
 *   V4 2026-02-29 → 非法，码 0117；2024-02-29 → 合法
 *   V5 2026-11-15 → 周内日 7（周日）
 * 红线自检 (Redline)    : R1 零全局变量表与外部变量引用 ｜ R2 零物理地址直写
 *                         R3 纯 IEC 61131-3 ｜ R4 域校验先判后算 + 除法除数恒为常量
 *                         R5 全变量中英双语同行注释 ｜ R6 CASE 含 ELSE 兜底（月份
 *                         查表用 CASE，非法月份走 ELSE）｜ R7 N/A（无实例调用）
 * 修订历史 (Revision)   :
 *   2026-11-15  v1.0.0  首版入库（Round 10 · Level 0 日历族回补）
 *============================================================================*)

FUNCTION FC_DL_WeekOfYearCalc : BOOL
VAR_INPUT
    nYear  : INT := 2026;   // 公历年，有效域 1970 到 2099 [年] / Calendar year, valid 1970 to 2099
    nMonth : INT := 1;      // 公历月，有效域 1 到 12 [月] / Calendar month, valid 1 to 12
    nDay   : INT := 1;      // 公历日，有效域 1 到该月天数 [日] / Day of month, valid 1 to month length
END_VAR
VAR_OUTPUT
    nIsoYear  : INT;        // ISO 周年，可能不等于 nYear（跨年归属所致）[年] / ISO week-numbering year, may differ from nYear
    nIsoWeek  : INT;        // ISO 周序号，1 到 53 [周] / ISO week number, 1 to 53
    nIsoDow   : INT;        // ISO 周内日，周一 = 1，周日 = 7 [1 到 7] / ISO day of week, Monday = 1, Sunday = 7
    nWeek53En : BOOL;       // 该 ISO 周年是否含第 53 周（长年判据）[布尔] / TRUE if that ISO year has week 53
    uErrorId  : UDINT;      // 事件码，0 = 无事件 / Event code, 0 = no event
END_VAR
VAR
    bLeapYear   : BOOL;     // 输入年是否闰年 [-] / TRUE if the input year is a leap year
    bLeapIso    : BOOL;     // ISO 周年是否闰年（长年判定用）[-] / TRUE if the ISO year is a leap year
    bPending    : BOOL;     // 周号待定标志（周四落到上一年时为 TRUE）[-] / TRUE when the week number must be resolved after the long-year test
    nMonthLen   : INT;      // 当月天数，随闰年调整 [日] / Length of the input month in days
    nDaysBefore : INT;      // 当月起点的年内序日偏移（不含当月 1 日）[日] / Day offset of the month start
    nDoy        : INT;      // 当日的年内序日，1 起 [日] / Day of year, 1-based
    nDaysInYear : INT;      // 输入年的总天数，365 或 366 [日] / Total days of the input year
    nThursday   : INT;      // 本周周四的年内序日，可能小于 1 或超过当年天数 [日] / Day of year of the Thursday of this week
    nZYear      : INT;      // Zeller 折算用年份（1 月 2 月取上一年）[年] / Year used by the Zeller term, shifted for January and February
    nZMonth     : INT;      // Zeller 折算用月份（1 月 2 月取 13 月 14 月）[月] / Month used by the Zeller term, shifted to 13 and 14
    nZCentury   : INT;      // Zeller 世纪项 J = 年 除以 100 [世纪] / Zeller century term J
    nZYearInC   : INT;      // Zeller 年内项 K = 年 对 100 取模 [年] / Zeller year-in-century term K
    nZMonthTerm : INT;      // Zeller 月份项，floor(13 乘 (月 加 1) 除以 5) [-] / Zeller month term
    nZSum       : INT;      // Zeller 求和中间量，域内不溢出 [-] / Zeller sum temporaries
    nZWeekday   : INT;      // Zeller 结果，0 = 周六，1 = 周日，2 = 周一，6 = 周五 [-] / Zeller weekday, 0 = Saturday
    nJan1IsoDow : INT;      // ISO 周年 1 月 1 日的 ISO 周内日 [1 到 7] / ISO weekday of January 1st of the ISO year
END_VAR
VAR CONSTANT
    DL_YEAR_MIN  : INT := 1970;   // 可算年下限 [年] / Lowest computable year
    DL_YEAR_MAX  : INT := 2099;   // 可算年上限 [年] / Highest computable year
    DL_WEEK_DAYS : INT := 7;      // 每周天数 [日] / Days per week
    DL_THU_KEY   : INT := 4;      // 周四的 ISO 周内日编号，周四归属法基准 [-] / ISO weekday index of Thursday
    DL_MONTH_MIN : INT := 1;      // 月份下限 [月] / Lowest month index
    DL_MONTH_MAX : INT := 12;     // 月份上限 [月] / Highest month index
    DL_DAY_MIN   : INT := 1;      // 日起点，0 与负数一律非法 [日] / Lowest day index
    DL_DAYS_COMMON : INT := 365;  // 平年天数 [日] / Days in a common year
    DL_DAYS_LEAP   : INT := 366;  // 闰年天数 [日] / Days in a leap year
    DL_WEEK_LAST   : INT := 52;   // 短年最后一周号 [周] / Last week number of a short ISO year
    DL_WEEK_LAST53 : INT := 53;   // 长年最后一周号 [周] / Last week number of a long ISO year
END_VAR

(*------------------------------------------------------------------------------
 * 段 1｜输出与返回值预置：任何早退路径下输出必须为确定的 0
 *      Pre-set outputs and return value: deterministic zeros on early exit
 *-----------------------------------------------------------------------------*)
FC_DL_WeekOfYearCalc := FALSE;
nIsoYear  := 0;
nIsoWeek  := 0;
nIsoDow   := 0;
nWeek53En := FALSE;
uErrorId  := 16#0000_0000;
bPending  := FALSE;

(*------------------------------------------------------------------------------
 * 段 2｜年份域校验（边界 B1）：早退，绝不带着非法年进入后续整除
 *      Year bounds check (boundary B1): early return before any integer division
 *-----------------------------------------------------------------------------*)
IF (nYear < DL_YEAR_MIN) OR (nYear > DL_YEAR_MAX) THEN
    uErrorId := 16#0001_0116;   // 年份越界，输出全 0
    RETURN;
END_IF

(*------------------------------------------------------------------------------
 * 段 3｜闰年判定：四年一闰、百年不闰、四百年再闰
 *      Leap year test: divisible by 4, not by 100, unless divisible by 400
 *-----------------------------------------------------------------------------*)
IF ((nYear MOD 4) = 0) AND (((nYear MOD 100) <> 0) OR ((nYear MOD 400) = 0)) THEN
    bLeapYear   := TRUE;
    nDaysInYear := DL_DAYS_LEAP;
ELSE
    bLeapYear   := FALSE;
    nDaysInYear := DL_DAYS_COMMON;
END_IF

(*------------------------------------------------------------------------------
 * 段 4｜月份天数与月首偏移查表（边界 B2）：CASE 带 ELSE 兜底，非法月份直接拒绝
 *      Month length and month-start offset lookup with an ELSE fallback branch
 *      用 CASE 而非数组常量，是为了让非法月份在 ELSE 里被显式拦下
 *-----------------------------------------------------------------------------*)
CASE nMonth OF
    1:
        nMonthLen   := 31;
        nDaysBefore := 0;
    2:
        nDaysBefore := 31;
        IF bLeapYear THEN
            nMonthLen := 29;     // 闰年 2 月 29 天
        ELSE
            nMonthLen := 28;     // 平年 2 月 28 天
        END_IF
    3:
        nMonthLen   := 31;
        nDaysBefore := 59;
        IF bLeapYear THEN
            nDaysBefore := 60;   // 闰年 3 月前多一天
        END_IF
    4:
        nMonthLen   := 30;
        nDaysBefore := 90;
        IF bLeapYear THEN
            nDaysBefore := 91;
        END_IF
    5:
        nMonthLen   := 31;
        nDaysBefore := 120;
        IF bLeapYear THEN
            nDaysBefore := 121;
        END_IF
    6:
        nMonthLen   := 30;
        nDaysBefore := 151;
        IF bLeapYear THEN
            nDaysBefore := 152;
        END_IF
    7:
        nMonthLen   := 31;
        nDaysBefore := 181;
        IF bLeapYear THEN
            nDaysBefore := 182;
        END_IF
    8:
        nMonthLen   := 31;
        nDaysBefore := 212;
        IF bLeapYear THEN
            nDaysBefore := 213;
        END_IF
    9:
        nMonthLen   := 30;
        nDaysBefore := 243;
        IF bLeapYear THEN
            nDaysBefore := 244;
        END_IF
    10:
        nMonthLen   := 31;
        nDaysBefore := 273;
        IF bLeapYear THEN
            nDaysBefore := 274;
        END_IF
    11:
        nMonthLen   := 30;
        nDaysBefore := 304;
        IF bLeapYear THEN
            nDaysBefore := 305;
        END_IF
    12:
        nMonthLen   := 31;
        nDaysBefore := 334;
        IF bLeapYear THEN
            nDaysBefore := 335;
        END_IF
    ELSE
        nMonthLen   := 0;        // 非法月份：不做任何推算
        nDaysBefore := 0;
        uErrorId    := 16#0001_0117;
        RETURN;
END_CASE

(*------------------------------------------------------------------------------
 * 段 5｜日期域校验（边界 B3）：日必须落在 1 到当月天数之间
 *      Day bounds check (boundary B3): day must be within the month length
 *-----------------------------------------------------------------------------*)
IF (nDay < DL_DAY_MIN) OR (nDay > nMonthLen) THEN
    uErrorId := 16#0001_0117;   // 日非法（含平年 2 月 29 日）
    RETURN;
END_IF

(*------------------------------------------------------------------------------
 * 段 6｜年内序日：月首偏移加当日，1 起
 *      Day of year: month-start offset plus the day, 1-based
 *-----------------------------------------------------------------------------*)
nDoy := nDaysBefore + nDay;

(*------------------------------------------------------------------------------
 * 段 7｜星期几（Zeller 同余重排）：1 月 2 月折算为上年的 13 月 14 月
 *      Weekday via a Zeller rearrangement: January and February shift to 13 and 14
 *      结果 0 = 周六，1 = 周日，2 = 周一，3 = 周二，4 = 周三，5 = 周四，6 = 周五
 *      再折算为 ISO 周内日：周一 1，周日 7，公式为 ((h 加 5) 对 7 取模) 加 1
 *-----------------------------------------------------------------------------*)
IF nMonth <= 2 THEN
    nZYear  := nYear - 1;       // 1 月 2 月归属上一年
    nZMonth := nMonth + 12;     // 1 月 改为 13 月，2 月 改为 14 月
ELSE
    nZYear  := nYear;
    nZMonth := nMonth;
END_IF

nZCentury   := nZYear / 100;                          // 世纪项 J
nZYearInC   := nZYear MOD 100;                        // 年内项 K
nZMonthTerm := (13 * (nZMonth + 1)) / 5;              // 月份项，整除向下取整
nZSum       := nDay + nZMonthTerm + nZYearInC
               + (nZYearInC / 4) + (nZCentury / 4) + (5 * nZCentury);

nZWeekday := nZSum MOD DL_WEEK_DAYS;                  // 0 = 周六 起算
nIsoDow   := ((nZWeekday + 5) MOD DL_WEEK_DAYS) + 1;  // 折算为 ISO 周内日

(*------------------------------------------------------------------------------
 * 段 8｜周四归属法：本周周四落在哪一年，本周就归属哪一年
 *      Thursday-ownership rule: the ISO year is the year of this week's Thursday
 *-----------------------------------------------------------------------------*)
nThursday := nDoy + (DL_THU_KEY - nIsoDow);   // 本周周四的年内序日，可为 0 或超过当年天数

IF nThursday < 1 THEN
    nIsoYear := nYear - 1;                    // 落在上一年：属上一年最后一周
    nIsoWeek := 0;                            // 周号待定（52 或 53），段 10 收口
    bPending := TRUE;
ELSIF nThursday > nDaysInYear THEN
    nIsoYear := nYear + 1;                    // 落在次年：属次年第 1 周
    nIsoWeek := 1;
ELSE
    nIsoYear := nYear;                        // 落在本年：正常整除求周号
    nIsoWeek := ((nThursday - 1) / DL_WEEK_DAYS) + 1;
END_IF

(*------------------------------------------------------------------------------
 * 段 9｜长年判定：ISO 周年 1 月 1 日为周四，或闰年且 1 月 1 日为周三
 *      Long-year test: January 1st is a Thursday, or a leap year starting on Wednesday
 *      长年含第 53 周；短年至第 52 周
 *-----------------------------------------------------------------------------*)
IF ((nIsoYear MOD 4) = 0) AND (((nIsoYear MOD 100) <> 0) OR ((nIsoYear MOD 400) = 0)) THEN
    bLeapIso := TRUE;
ELSE
    bLeapIso := FALSE;
END_IF

(* 复用同一套 Zeller 重排式，仅把入参固定为 ISO 周年的 1 月 1 日 *)
nZYear      := nIsoYear - 1;                    // 1 月 归属上一年
nZCentury   := nZYear / 100;
nZYearInC   := nZYear MOD 100;
nZMonthTerm := (13 * 14) / 5;                   // 14 月 的月份项，常量 36
nZSum       := 1 + nZMonthTerm + nZYearInC
               + (nZYearInC / 4) + (nZCentury / 4) + (5 * nZCentury);
nZWeekday   := nZSum MOD DL_WEEK_DAYS;
nJan1IsoDow := ((nZWeekday + 5) MOD DL_WEEK_DAYS) + 1;

IF (nJan1IsoDow = DL_THU_KEY) OR (bLeapIso AND (nJan1IsoDow = (DL_THU_KEY - 1))) THEN
    nWeek53En := TRUE;                          // 长年，含第 53 周
ELSE
    nWeek53En := FALSE;                         // 短年，最后一周为第 52 周
END_IF

(*------------------------------------------------------------------------------
 * 段 10｜跨年周号收口：周四落上一年时，按上一年是长年还是短年取 53 或 52
 *      Pending week resolution: 53 for a long ISO year, 52 for a short one
 *-----------------------------------------------------------------------------*)
IF bPending THEN
    IF nWeek53En THEN
        nIsoWeek := DL_WEEK_LAST53;
    ELSE
        nIsoWeek := DL_WEEK_LAST;
    END_IF
END_IF

(*------------------------------------------------------------------------------
 * 段 11｜返回值收口：三段输出均已赋值，标记计算成功
 *      Close-out: all three outputs assigned, flag success
 *-----------------------------------------------------------------------------*)
FC_DL_WeekOfYearCalc := TRUE;
END_FUNCTION

(* ---- FC_DL_WordsToDword.st ---- *)
(*==============================================================================
 * 名称 : FC_DL_WordsToDword —— 两个 WORD 合成 DWORD（显式高低序参数）
 * 分类 / 前缀 / 版本 : DL_Base / FC_DL_ / 1.0.0
 * 溯源 : 开源语义参考（OSCAT/AixOCAT 族，MIT）或 clean-room IEC 实现，未复制源码
 * 平台 : 纯 IEC 61131-3
 * 功能说明 : 将两个 16 位 WORD 合成为 32 位 DWORD：bFirstIsHigh=TRUE 时 wFirst
 *            为高字、wSecond 为低字；FALSE 时角色对调。
 *            合成全程数值语义（WORD_TO_DWORD + SHL/OR），不触碰内存序。
 *            边界处理：两字覆盖完整 32 位，无溢出；与 FC_DL_DwordToWords 互为
 *            逆运算（同参数口径下往返一致）。
 * 错误码 : 无故障路径（全值域合法的纯合成），eErr 恒 0，bValid 恒 TRUE；
 *          16#0001_1A0B 为本件预留码位，当前实现不发出
 * 状态机 : R6 标注 N/A（纯函数无顺序状态，以本节替代 ELSE 兜底）
 * 红线 : R1/R2/R3 ✓ 零全局/零IO/纯IEC ｜ R4 ✓ 移位量=16 ｜ R10 ✓ 标准转换 ｜ R11 ✓ 分号收尾 ｜ R15 ✓ 无保留字撞名
 * 修订记录 : 2026-11-23 v1.0.0 首次入库（R76）
 *============================================================================*)
FUNCTION FC_DL_WordsToDword : DWORD
VAR_INPUT
    wFirst      : WORD;    // 首个输入字 [位域] / first input word
    wSecond     : WORD;    // 第二个输入字 [位域] / second input word
    bFirstIsHigh: BOOL;    // TRUE=wFirst 为高字 / TRUE when wFirst is the high word
END_VAR
VAR_OUTPUT
    eErr   : UDINT;    // 故障码，0=正常（本件无故障路径）/ error code, 0=ok (no fault path)
    bError : BOOL;     // 故障标志，恒 FALSE / error flag, always FALSE
    bValid : BOOL;     // TRUE=返回值可用，恒 TRUE / TRUE when return value is usable
END_VAR
VAR
    _wHi : WORD;       // 判定后的高字 [位域] / resolved high word
    _wLo : WORD;       // 判定后的低字 [位域] / resolved low word
END_VAR

eErr   := 16#0000_0000;                      // 故障码清零 / clear error code
bError := FALSE;                             // 故障标志清零 / clear error flag
bValid := TRUE;                              // 本件全值域合法，恒可用 / always valid

IF bFirstIsHigh THEN                         // wFirst 为高字 / wFirst is high
    _wHi := wFirst;                          // 取 wFirst 为高字 / take wFirst as high
    _wLo := wSecond;                         // 取 wSecond 为低字 / take wSecond as low
ELSE                                         // wSecond 为高字 / wSecond is high
    _wHi := wSecond;                         // 取 wSecond 为高字 / take wSecond as high
    _wLo := wFirst;                          // 取 wFirst 为低字 / take wFirst as low
END_IF

FC_DL_WordsToDword := SHL(WORD_TO_DWORD(_wHi), 16) OR WORD_TO_DWORD(_wLo);    // 高字左移 16 位后并入低字（移位量 16<32 安全）/ compose

END_FUNCTION

(* ---- FC_DL_WorkdayCalendarCalc.st ---- *)
// FC_DL_WorkdayCalendarCalc v1.0.0
// 开源溯源：self-cleanroom / 公历算法（Fliegel-Van Flandern 公开公式）
(*
  道莅工业代码库 | DL_Base | FC_DL_WorkdayCalendarCalc
  版本: 1.0.0 | 日期: 2026-11-23 | 轮次: R75
  功能: 日期区间工作日计数（周一~周五，剔除内嵌节假日表命中项）；
        儒略日数算法取星期，整周×5 + 余数逐日扫描，节假日逐项扣减
  邻件关系: 与 WeekNumIsoCalc / DateDiffDays / DayOfWeekCalc 同族 —— 差异点：
            周号件算 ISO 周、差值件算自然日差，本件算工作日净计数（含
            节假日剔除），星期口径经 JDN MOD 7 自证（2026-11-23 周一 = 0）
  日期契约: 入参为 DINT 型 yyyymmdd 十进制编码（如 20261123）；
            节假日表 aHoliday 同口径，nHolidayCnt 个有效（0..16）
*)
FUNCTION FC_DL_WorkdayCalendarCalc : DINT
VAR_INPUT
    dStart       : DINT;                          // 起始日期 [yyyymmdd 编码] / Start date as yyyymmdd
    dEnd         : DINT;                          // 结束日期（含当日）[yyyymmdd] / End date inclusive, as yyyymmdd
    aHoliday     : ARRAY[1..16] OF DINT;          // 节假日表 [yyyymmdd 编码] / Holiday table as yyyymmdd
    nHolidayCnt  : INT;                           // 节假日有效个数 [个]，域 0..16 / Valid holiday count
END_VAR
VAR_OUTPUT
    bValid       : BOOL;                          // 结果有效回执 [-] / Result validity receipt
    nWorkdays    : DINT;                          // 工作日计数 [天] / Workday count [days]
    uErrorId     : UDINT;                         // 事件码，0 = 无事件；16#0002_2301 = 日期非法 / Event code
END_VAR
VAR
    nSx          : DINT;                          // 起始年 [年] / Start year
    nSm          : DINT;                          // 起始月 [月] / Start month
    nSd          : DINT;                          // 起始日 [日] / Start day
    nEx          : DINT;                          // 结束年 [年] / End year
    nEm          : DINT;                          // 结束月 [月] / End month
    nEd          : DINT;                          // 结束日 [日] / End day
    nTmp         : DINT;                          // 交换/中间量 [—] / Swap temp
    nTotalDays   : DINT;                          // 区间自然日总数（含端点）[天] / Total days inclusive
    nJdnS        : DINT;                          // 起始儒略日数 [天] / Start JDN
    nFullWeeks   : DINT;                          // 整周数 [周] / Full weeks
    nRemain      : DINT;                          // 余数天数 [天] / Remainder days
    nCount       : DINT;                          // 工作日累计 [天] / Workday accumulator
    nDow         : DINT;                          // 星期（0=周一..6=周日）[1] / Day of week, 0=Mon..6=Sun
    nJdnCur      : DINT;                          // 余数段当前儒略日 [天] / Current JDN in remainder scan
    h            : INT;                           // 节假日表索引 [个] / Holiday table index
    dHol         : DINT;                          // 当前节假日 [yyyymmdd] / Current holiday
    nJdnHol      : DINT;                          // 节假日儒略日 [天] / Holiday JDN
    bHolInRange  : BOOL;                          // 节假日落在区间内 [-] / Holiday within range
END_VAR
VAR CONSTANT
    DL_WDC_JDN_EPOCH_OFF : DINT := 32075;         // Fliegel 公式尾部常数 [天] / Fliegel tail constant
END_VAR

// —— 段 0：全路径缺省 —— //
bValid := FALSE;                                     // 有效回执预清 / Validity preset
nWorkdays := 0;                                      // 计数缺省零 / Count default zero
uErrorId := 16#0000;                                 // 事件码预清 / Event code preset
FC_DL_WorkdayCalendarCalc := 0;                      // 返回值缺省零 / Return default zero

// —— 段 1：日期编码与区间闸（格式 + 序向） —— //
IF dStart > dEnd THEN                                // 起点晚于终点：交换（宽容序）/ Swap tolerant order
    nTmp := dStart;
    dStart := dEnd;
    dEnd := nTmp;
END_IF
nSx := dStart / 10000;                               // 年提取 [年] / Year extract
nSm := (dStart MOD 10000) / 100;                     // 月提取 [月] / Month extract
nSd := dStart MOD 100;                               // 日提取 [日] / Day extract
nEx := dEnd / 10000;
nEm := (dEnd MOD 10000) / 100;
nEd := dEnd MOD 100;
IF (nSm < 1) OR (nSm > 12) OR (nEm < 1) OR (nEm > 12)
   OR (nSd < 1) OR (nSd > 31) OR (nEd < 1) OR (nEd > 31) THEN   // 月日域闸 / Month and day domain gate
    uErrorId := 16#0002_2301;                        // 信息级：日期编码非法 / Info level: illegal date code
    RETURN;
END_IF
IF (nHolidayCnt < 0) OR (nHolidayCnt > 16) THEN      // 节假日计数域闸 / Holiday count gate
    uErrorId := 16#0002_2301;                        // 计数非法同码段 / Same code family
    RETURN;
END_IF

// —— 段 2：儒略日数（Fliegel-Van Flandern，整数除即 ST DIV 截断口径） —— //
nJdnS := (1461 * (nSx + 4800 + (nSm - 14) / 12)) / 4
         + (367 * (nSm - 2 - 12 * ((nSm - 14) / 12))) / 12
         - (3 * ((nSx + 4900 + (nSm - 14) / 12) / 100)) / 4
         + nSd - DL_WDC_JDN_EPOCH_OFF;               // 起始 JDN [天] / Start JDN
nTmp := (1461 * (nEx + 4800 + (nEm - 14) / 12)) / 4
        + (367 * (nEm - 2 - 12 * ((nEm - 14) / 12))) / 12
        - (3 * ((nEx + 4900 + (nEm - 14) / 12) / 100)) / 4
        + nEd - DL_WDC_JDN_EPOCH_OFF;                // 结束 JDN（复用暂存）/ End JDN
nTotalDays := nTmp - nJdnS + 1;                      // 含端点自然日 [天] / Inclusive day count

// —— 段 3：整周×5 工作日基数 —— //
nFullWeeks := nTotalDays / 7;                        // 整周数 [周] / Full weeks
nRemain := nTotalDays - nFullWeeks * 7;              // 余数天 [天] / Remainder days
nCount := nFullWeeks * 5;                            // 整周工作日基数 [天] / Full-week weekday base

// —— 段 4：余数段逐日扫描（起点 JDN 起，nRemain ≤ 6 循环有界） —— //
nJdnCur := nJdnS;                                    // 扫描游标 [天] / Scan cursor
FOR nTmp := 1 TO nRemain DO                           // 余数天逐日（≤6 次）/ Day scan, bounded
    nDow := (nJdnCur MOD 7);                         // 星期 0=周一..6=周日（自证：2026-11-23 JDN MOD 7 = 0 = 周一）/ Dow 0=Mon..6=Sun
    IF nDow <= 4 THEN                                // 周一~周五 / Monday to Friday
        nCount := nCount + 1;                        // 工作日累加 / Count workday
    END_IF
    nJdnCur := nJdnCur + 1;                          // 游标前进 / Advance cursor
END_FOR

// —— 段 5：节假日扣减（表内逐项：在区间内且为工作日则扣 1） —— //
FOR h := 1 TO nHolidayCnt DO                         // 逐节假日（h ≤ nHolidayCnt ≤ 16 判界安全）/ Per holiday, index safe
    dHol := aHoliday[h];                             // 取节假日编码 / Holiday code
    IF (dHol MOD 10000) / 100 >= 1 AND (dHol MOD 10000) / 100 <= 12 AND (dHol MOD 100 >= 1) AND (dHol MOD 100 <= 31) THEN
        nJdnHol := (1461 * (dHol / 10000 + 4800 + ((dHol MOD 10000) / 100 - 14) / 12)) / 4
                   + (367 * ((dHol MOD 10000) / 100 - 2 - 12 * (((dHol MOD 10000) / 100 - 14) / 12))) / 12
                   - (3 * ((dHol / 10000 + 4900 + ((dHol MOD 10000) / 100 - 14) / 12) / 100)) / 4
                   + (dHol MOD 100) - DL_WDC_JDN_EPOCH_OFF;   // 节假日 JDN [天] / Holiday JDN
        bHolInRange := (nJdnHol >= nJdnS) AND (nJdnHol <= nJdnS + nTotalDays - 1);   // 区间内判据 / In-range test
        IF bHolInRange THEN
            nDow := (nJdnHol MOD 7);                 // 节假日星期 [1] / Holiday dow
            IF nDow <= 4 THEN                        // 仅工作日节假日扣减（周末节假日已不在基数）/ Deduct only weekday holidays
                nCount := nCount - 1;                // 扣减 / Deduct
            END_IF
        END_IF
    END_IF
END_FOR

// —— 段 6：输出收口 —— //
IF nCount < 0 THEN
    nCount := 0;                                     // 负值兜底（防御）/ Negative guard
END_IF
nWorkdays := nCount;                                 // 计数输出 / Count output
bValid := TRUE;                                      // 有效回执 / Validity receipt
FC_DL_WorkdayCalendarCalc := nCount;                 // 返回值 = 工作日数 / Return equals count
END_FUNCTION

(* ---- FB_DL_AlarmFloodLimiter.st ---- *)
(*==============================================================================
 * 组件名称 (Component)  : FB_DL_AlarmFloodLimiter
 * 所属子库 (Sublibrary) : DL_Base
 * 当前版本 (Version)    : 1.0.0
 * 兼容性   (Platform)   : CODESYS 3.5+ / TwinCAT 3 / 汇川 InoProShop / 施耐德 Machine Expert
 *                         仅依赖 Standard.library（TON / R_TRIG），零厂商私有库
 * 功能描述 (Function)   : 报警泛滥抑制（ISA-18.2 泛滥抑制语义）。同源报警在一个分窗内
 *                         累计次数超过 nFloodLimit 即进入抑制态 bSuppressed；抑制期
 *                         tSuppressHold 内新报警不再上送（bPassThrough = FALSE），但抑制期
 *                         内到达的报警仍逐次计数，抑制结束时以 nSuppressedCount 一次性
 *                         给出该段台账（首末计数语义：进入抑制清零，抑制结束定稿）。
 *                         禁止抑制任何「安全类」来源：bSafetyCritical 为真时 bPassThrough
 *                         恒为真，且该类报警不进入泛滥计数（安全侧不可被闸掉，本件核心红线）。
 * 接口     (Interface)  : 输入 uAlarmSrc 来源号、bAlarmActive 报警有效位、bSafetyCritical
 *                         安全类标记、nFloodLimit 窗内同源次数上限、tWindow 分窗时长、
 *                         tSuppressHold 抑制保持时长、bReset 复位电平；输出 bPassThrough
 *                         上送许可、bSuppressed 抑制态、nSuppressedCount 抑制期计数台账、
 *                         nWindowCount 当前窗计数、eState / eCause / bError / nErrId。
 * 边界     (Boundary)   : ① 组态闸：nFloodLimit = 0 或 tWindow <= T#0S 或 tSuppressHold <= T#0S
 *                         → 故障锁存；② 分窗用 TON 自复位实现（IN := NOT tonWindow.Q，
 *                         R188），窗口边界由计时器自身产生，不依赖外部沿清零；
 *                         ③ **不使用数组环缓冲**，故本件无下标越界路径（派单「环缓冲下标先判
 *                         边界」条款在本件以「零数组」方式结构性满足）；
 *                         ④ TON 两枚 + R_TRIG 两枚段 0 无条件周期刷新；
 *                         ⑤ 故障相迁出唯一路径 = bReset 上升沿；⑥ 零全局耦合（无 GVL / 无物理地址）。
 * 解除式   (Release)    : bReset 上升沿 ∧ 组态合法 ∧ 抑制态已退出（NOT bSuppressed，当拍量，
 *                         R240 范式）。自证可满足（终审两式 1）：tonSuppress 的 IN 挂抑制态
 *                         本身，抑制态退出后 IN 落假、Q 必落假，且组态修正后闸即放开，无恒假因子。
 * 码表     (Codes)      : 16#0001_03EC 故障级：泛滥抑制器故障总码（组态非法 / 非法相位），
 *                         锁存至 bReset 上升沿，归因由 eCause 承载（R190 单件单总码）；
 *                         16#0001_04AF 信息级：抑制段结束台账（抑制保持期到，nSuppressedCount 定稿）。
 *                         加码反证（R90）：抑制段结束是一个不改变 bSuppressed 终值的「已发生事实」，
 *                         其唯一可观测证据是抑制期累计数，而该数在抑制结束后与抑制前的
 *                         nWindowCount 无任何可分辨关系，故须立一码留痕。
 *                         码段说明：0001 段故障子带 03xx / 信息子带 04xx，本件取 03EC / 04AF
 *                         （源码实扫该两槽为空，续接同子带已用最大值，未回填碎片孔洞）。
 * 开源溯源 (Origin)     : 道莅自研 clean-room（参考 ISA-18.2 报警生命周期分类与参数域，
 *                         零代码行复制；t2-8-isa182 族）
 * 修订历史 (Revision)   : 2026-11-19  v1.0.0  R45 首版（批次 1 · 序号 3）
 *==============================================================================*)

TYPE E_DL_AflState :
(
    eIdle  := 0,     // 窗内无报警流量，等待首个报警 / Idle, no alarm traffic in window
    eRun   := 10,    // 计数/抑制运行 / Counting or suppressing
    eFault := 90     // 故障锁存相 / Fault latched phase
);
END_TYPE

TYPE E_DL_AflCause :
(
    eNone       := 0,   // 无故障成因 / No cause
    eCfgIllegal := 1    // 组态非法 / Illegal configuration
);
END_TYPE

FUNCTION_BLOCK FB_DL_AlarmFloodLimiter
VAR_INPUT
    uAlarmSrc       : UINT := 0;              // 报警来源号，同号视为同源 [号] / Alarm source id, same id means same source
    bAlarmActive    : BOOL := FALSE;          // 报警有效位（电平），上升沿计入一次 [次] / Alarm active level, rising edge counts once
    bSafetyCritical : BOOL := FALSE;          // 安全类来源标记，TRUE 时永不被抑制 [-] / Safety-critical source, never suppressed when TRUE
    nFloodLimit     : UDINT := 10;            // 窗内同源次数上限，域 > 0 [次] / Same-source count limit in window, domain > 0
    tWindow         : TIME := T#10S;          // 分窗时长，域 > T#0S [ms] / Window duration, domain > T#0S
    tSuppressHold   : TIME := T#60S;          // 抑制保持时长，域 > T#0S [ms] / Suppression hold duration
    bReset          : BOOL := FALSE;          // 复位命令，上升沿清故障 [-] / Reset command, rising edge clears fault
END_VAR
VAR_OUTPUT
    bPassThrough      : BOOL;                 // 上送许可，TRUE = 允许报警上送 [-] / Pass-through permit for alarm upload
    bSuppressed       : BOOL;                 // 抑制态镜像 [-] / Suppression state mirror
    nSuppressedCount  : UDINT;                // 抑制期计数台账（锁存量，抑制结束定稿） [次] / Suppressed count ledger, latched
    nWindowCount      : UDINT;                // 当前分窗内同源计数 [次] / Same-source count in current window
    eState            : E_DL_AflState;        // 状态出口，段 6 单点映射 / State outlet
    eCause            : E_DL_AflCause;        // 故障成因出口（R190 归因唯一） / Fault cause outlet
    bError            : BOOL;                 // 故障锁存标志 [-] / Fault latch flag
    nErrId            : UDINT;                // 事件码，0 = 无事件 / Event code, 0 = no event
END_VAR
VAR
    _eState           : E_DL_AflState := E_DL_AflState.eIdle;   // 内部相位（CASE 唯一写入目标） / Internal phase
    _eCause           : E_DL_AflCause := E_DL_AflCause.eNone;   // 故障成因锁存（锁存量） / Latched cause
    tonWindow         : TON;                  // 分窗计时（自复位），段 0 无条件调用 / Window timer, self-resetting
    tonSuppress       : TON;                  // 抑制保持计时，段 0 无条件调用 / Suppression hold timer
    rtAlarm           : R_TRIG;               // 报警上升沿实例，段 0 无条件调用 / Alarm rising edge
    rtReset           : R_TRIG;               // 复位沿实例，段 0 无条件调用 / Reset edge
    _bSuppressed      : BOOL;                 // 抑制态（锁存量） / Suppression state, latched
    _nWindowCount     : UDINT;                // 窗内同源计数（锁存量，唯一写入点） [次] / Window count, single write point
    _nSuppCount       : UDINT;                // 抑制期累计计数（锁存量，唯一写入点） [次] / Suppressed cumulative count, single write point
    _uSrcLast         : UINT;                 // 上一报警来源号（窗内归属判定） [号] / Last alarm source id for window attribution
    _bCfgBad          : BOOL;                 // 组态非法当拍量 [-] / Illegal configuration
    _bFault           : BOOL;                 // 故障锁存位（锁存量） / Latched fault bit
    _uFault           : UDINT;                // 故障码锁存（锁存量） / Latched fault code
    _uInfo            : UDINT;                // 信息码，每拍重算 / Info code, recomputed each scan
END_VAR
VAR CONSTANT
    DL_COUNT_MAX : UDINT := 16#FFFF_FFFE;     // 计数饱和上限，留加 1 裕度防溢出 [次] / Count saturation limit with increment margin [count]
END_VAR

(* —— 段 0：当拍量派生 + 定时器与沿实例无条件周期刷新 —— *)
_bCfgBad := (nFloodLimit = 0) OR (tWindow <= T#0S) OR (tSuppressHold <= T#0S);  // 组态非法当拍量 / Illegal configuration
rtAlarm(CLK := bAlarmActive);                                                   // 报警沿，每拍必调（R228A） / Alarm edge, called every scan
rtReset(CLK := bReset);                                                         // 复位沿，每拍必调 / Reset edge, called every scan
tonWindow(IN := NOT tonWindow.Q, PT := tWindow);                                // 分窗计时自复位（R188） / Self-resetting window timer
tonSuppress(IN := _bSuppressed, PT := tSuppressHold);                           // 抑制保持计时，IN 挂抑制态 / Suppression hold timer gated by state

(* —— 段 1：单拍量预清零（锁存量不入清单，R107） —— *)
_uInfo           := 16#0000_0000;        // 信息码每拍重算 / Info recomputed every scan
nErrId           := 16#0000_0000;        // 事件码缺省无事件 / Event code default none
bError           := FALSE;               // 故障标志每拍预清，故障分支同拍置位（R45 配对） / Flag preset
bPassThrough     := TRUE;                // 上送许可缺省允许（安全侧优先） / Pass-through defaults to TRUE, safe side
bSuppressed      := _bSuppressed;        // 抑制态镜像（名实同源） / Suppression mirror
nSuppressedCount := _nSuppCount;         // 抑制台账镜像（锁存量回放） / Suppressed ledger mirror
nWindowCount     := _nWindowCount;       // 窗计数镜像（锁存量回放） / Window count mirror

(* —— 段 2：复位沿 + 组态域闸 —— *)
IF rtReset.Q THEN                                                        // 当拍复位沿 / current-scan reset edge
    _bFault := FALSE;                                                    // 清故障锁存位（锁存量） / Clear fault latch
    _uFault := 16#0000_0000;                                             // 清故障锁存码（锁存量） / Clear latched code
    _eCause := E_DL_AflCause.eNone;                                      // 清成因（锁存量） / Clear latched cause
    IF _eState = E_DL_AflState.eFault THEN
        _eState := E_DL_AflState.eIdle;                                  // 故障相迁出唯一路径 / Sole exit from fault phase
    END_IF
END_IF
IF _bCfgBad THEN                                                         // 组态域闸 / Configuration gate
    _uFault := 16#0001_03EC;                                             // 故障级：泛滥抑制器故障总码 / Fault-level: limiter fault code
    _bFault := TRUE;
    bError  := TRUE;                                                     // 故障标志同拍置位（R45 配对） / Error flag set same scan
    _eCause := E_DL_AflCause.eCfgIllegal;                                // 归因：组态非法 / Cause: illegal configuration
END_IF

(* —— 段 3：分窗边界 / 泛滥计数 / 抑制保持 —— *)
IF tonWindow.Q THEN                                                      // 窗口边界（单拍事件，自复位产生） / Window boundary, single scan
    _nWindowCount := 0;                                                  // 新窗计数清零（窗内量唯一重置点） / Reset window count at boundary
    _uSrcLast := 0;                                                      // 新窗来源归属清零 / Reset source attribution
END_IF
IF (NOT _bFault) AND rtAlarm.Q AND (NOT bSafetyCritical) THEN            // 安全类不入泛滥计数（红线） / Safety alarms excluded from flood counting
    IF (NOT _bSuppressed) THEN
        IF uAlarmSrc = _uSrcLast THEN                                    // 同源（整数判等合法） / Same source, integer equality is legal
            IF _nWindowCount < DL_COUNT_MAX THEN
                _nWindowCount := _nWindowCount + 1;                      // 同源计数递增 / Same-source increment
            END_IF
        ELSE
            _uSrcLast := uAlarmSrc;                                      // 换源重开计数 / New source restarts counting
            _nWindowCount := 1;
        END_IF
        IF _nWindowCount > nFloodLimit THEN                              // 超限进抑制 / Over limit enters suppression
            _bSuppressed := TRUE;                                        // 抑制态置位（锁存量） / Suppression latched
            _nSuppCount := 0;                                            // 抑制期台账清零（进入唯一重置点） / Ledger reset at entry
        END_IF
    ELSE
        IF _nSuppCount < DL_COUNT_MAX THEN
            _nSuppCount := _nSuppCount + 1;                              // 抑制期仍继续计数 / Counting continues while suppressed
        END_IF
    END_IF
END_IF
IF _bSuppressed AND tonSuppress.Q THEN                                   // 抑制保持期到 / Suppression hold elapsed
    _bSuppressed := FALSE;                                               // 退出抑制（锁存量） / Exit suppression
    _uInfo := 16#0001_04AF;                                              // 信息级：抑制段结束台账 / Info: suppression segment closed
    _nWindowCount := 0;                                                  // 抑制结束重开窗计数 / Restart window counting
    _uSrcLast := 0;                                                      // 抑制结束清来源归属 / Clear source attribution
END_IF

(* —— 段 4：故障解除式（R240 全当拍量） —— *)
IF rtReset.Q AND (NOT _bCfgBad) AND (NOT _bSuppressed) THEN
    _bFault := FALSE;                                                    // 清故障锁存位（锁存量） / Clear fault latch
    _uFault := 16#0000_0000;                                             // 清故障锁存码（锁存量） / Clear latched code
    _eCause := E_DL_AflCause.eNone;                                      // 清成因（锁存量） / Clear latched cause
END_IF

(* —— 段 4A：故障锁存相位迁移闸 —— *)
IF _bFault AND (_eState <> E_DL_AflState.eFault) THEN
    _eState := E_DL_AflState.eFault;                                     // 锁存即入故障相 / Latch enters fault phase
END_IF

(* —— 段 5：相位机（ENUM 全成员显式标签 + ELSE 兜底，R128） —— *)
CASE _eState OF

E_DL_AflState.eIdle:
    IF (_nWindowCount > 0) OR _bSuppressed THEN                           // 出口 1：窗内有流量或抑制中 / Traffic present or suppressing
        _eState := E_DL_AflState.eRun;
    ELSIF _bFault THEN                                                    // 出口 2：故障锁存 / Fault latched
        _eState := E_DL_AflState.eFault;
    END_IF

E_DL_AflState.eRun:
    IF (_nWindowCount = 0) AND (NOT _bSuppressed) THEN                    // 出口 1：窗空且未抑制 / Empty window, not suppressing
        _eState := E_DL_AflState.eIdle;
    ELSIF _bFault THEN                                                    // 出口 2：故障锁存 / Fault latched
        _eState := E_DL_AflState.eFault;
    END_IF

E_DL_AflState.eFault:
    ;                                                                      // 故障相：仅段 4 复位沿可迁出 / Only the reset edge leaves this phase

ELSE
    _uFault := 16#0001_03EC;                                              // 故障级：非法相位兜底（归并总码） / Illegal-phase fallback
    _bFault := TRUE;
    bError  := TRUE;
    _eCause := E_DL_AflCause.eCfgIllegal;                                 // 归因：相位非法归并组态 / Cause: phase illegal
    _eState := E_DL_AflState.eFault;

END_CASE

(* —— 段 6：出口单点映射（名实同源；锁存码回放；安全侧钳位） —— *)
IF bSafetyCritical OR _bFault THEN
    bPassThrough := TRUE;                                                 // 安全类 / 故障相恒放行（核心红线，不掩盖报警） / Always pass for safety sources and in fault
ELSIF _bSuppressed THEN
    bPassThrough := FALSE;                                                // 抑制期闸掉（仅非安全类、无故障） / Gated while suppressing
ELSE
    bPassThrough := TRUE;                                                 // 默认放行 / Default permit
END_IF
IF _bFault THEN
    nErrId := _uFault;                                                    // 故障锁存码回放 / Replay latched fault code
ELSE
    nErrId := _uInfo;                                                     // 信息码 / Info code
END_IF
bError := _bFault;                                                        // 故障标志与锁存同源（名实双出口，R191） / Flag from latch
eState := _eState;                                                        // 状态出口 / State outlet
eCause := _eCause;                                                        // 成因出口 / Cause outlet

END_FUNCTION_BLOCK

(* ---- FB_DL_AlarmManager.st ---- *)
(*==============================================================================
 * 组件名称 (Component)  : FB_DL_AlarmManager
 * 所属子库 (Sublibrary) : DL_Base
 * 当前版本 (Version)    : 1.0.0
 * 兼容性   (Platform)   : CODESYS 3.5 / TwinCAT 3 / 汇川 InoProShop / Machine Expert
 *                         仅依赖 Standard.library（R_TRIG）+ 本库位打包构件
 * 功能描述 (Function)   : 16 通道报警优先级仲裁器。通道可配停机级 / 警告级 / 提示级 /
 *                         禁用四档；输出激活报警字、激活通道数、停机联锁位、
 *                         首出通道索引与当前最高优先级通道索引。
 *                         首出采用"先到先得"序号仲裁：每通道在激活沿取一个全局递增序号，
 *                         首出即序号最小者，与通道物理位置无关，避免低位通道永远抢先。
 *                         确认只清除首出锁存、不清除激活态——激活 / 已确认 / 首出锁存
 *                         三个信号正交输出，这是报警管理的基本纪律。
 *                         只做仲裁与锁存，不做事件历史与抑制管理（属上位机职责）。
 * 开源溯源 (Origin)     : 原创实现。优先级分级、首出锁存、确认三态分离等概念
 *                         参照 ISA-18.2 报警管理方法论的公开描述；代码为本库独立重构，
 *                         未复制任何源码。
 * 本文件内含       : FB    FB_DL_AlarmManager（单 POU，无配套类型）
 * 依赖     (Depends)    : FC_DL_PackBitsToWord（首轮 #6，报警字打包）
 *                         Standard.library: R_TRIG
 * 红线自检 (Redline)    : R1 ✓ 禁用全局存储与物理寻址 ｜ R2 ✓ 无地址直写
 *                         R3 ✓ 纯 IEC 61131-3 ｜ R4 ✓ 数组双检 + 序号饱和 + 优先级钳位
 *                         R5 ✓ 全变量中英双语同行注释 ｜ R6 N/A（仲裁为每周期全量重算，
 *                            无跨周期状态转移，故以本节说明替代 ELSE 兜底）
 *                         R7 ✓ R_TRIG 主体最前部无条件刷新 ｜ R8 ✓ 通道数与优先级全常量化
 *
 * 【首出语义：电平敏感 / First-out is level-sensitive（决策 D-R2-04）】
 *   输入即"报警态信号"（TRUE = 正在报警）。冷启动时已处于报警态的通道
 *   会在首扫按扫描顺序依次取号，因而谁先被扫到谁就是首出——
 *   这是电平敏感方案的固有行为，手册必须写明；需要"相对已知良好起点"判定
 *   的场合应由调用方在输入侧做沿处理。
 *
 * 【确认语义 / Acknowledge semantics（决策 D-R2-07）】
 *   确认沿只推进序号水位并清首出锁存，不改变任何通道的激活态。
 *   确认后若有更新的报警，按序号顺序自动补位成为新首出；
 *   已确认但仍在报警的通道不会再次成为首出，直到它消失后重新激活。
 *
 * 【使能恢复语义 / Re-enable semantics（决策 P6）】
 *   禁用会清空序号表与全部输出，重新使能视同冷启动重扫，
 *   避免"禁用期间积压的报警在恢复瞬间集中爆发、首出指向历史事件"的混淆。
 *
 * 修订历史 (Revision)   :
 *   2026-11-14  v1.0.0  首版入库（Phase 1 第二轮 · Level 0 批次 D）
 *============================================================================*)
FUNCTION_BLOCK FB_DL_AlarmManager
VAR_INPUT
    abAlarmActive : ARRAY[0..15] OF BOOL;   // 16 路报警激活态，电平敏感 / 16 alarm active levels, level-sensitive
    auPriority    : ARRAY[0..15] OF USINT;  // 通道优先级，0=禁用 1=停机 2=警告 3=提示 / Channel priority
    bAck          : BOOL;                   // 上升沿确认：清除首出锁存 / Rising edge: acknowledge the first-out latch
    bEnable       : BOOL := TRUE;           // 使能，FALSE 时全部输出清零 / Enable, FALSE clears every output
END_VAR
VAR_OUTPUT
    uAlarmWord    : WORD;    // 激活报警位图，bit0 = 通道 0，仅含启用通道 / Active bitmap, bit0 = channel 0, enabled only
    uActiveCount  : USINT;   // 激活通道数 [个]，值域 0..16 / Active channel count [count], range 0..16
    bAnyActive    : BOOL;    // 存在任意激活报警 / Any alarm active
    bShutdown     : BOOL;    // 存在停机级激活报警（联锁用）/ Any stop-level alarm active, for interlocking
    nFirstOutIdx  : INT;     // 首出通道索引，-1 = 无 / First-out channel index, -1 = none
    bFirstOutAck  : BOOL;    // 首出已确认标志 / First-out acknowledged flag
    nTopPrioIdx   : INT;     // 当前最高优先级激活通道（同级先到先得），-1 = 无 / Top-priority active channel, -1 = none
    uErrorId      : UDINT;   // 故障码，0 = 无故障 / Error code, 0 = no error
END_VAR
VAR
    auSeqNo       : ARRAY[0..15] OF UDINT;  // 通道激活序号，0 = 从未激活 / Activation sequence number, 0 = never activated
    auPrioEff     : ARRAY[0..15] OF USINT;  // 钳位后的通道优先级 / Clamped channel priority
    abPackSrc     : ARRAY[0..15] OF BOOL;   // 打包源（禁用通道置 FALSE）/ Packing source, disabled channels forced FALSE
    uSeqNext      : UDINT;                  // 全局递增序号发生器 / Global sequence generator
    uAckSeq       : UDINT;                  // 最近一次确认时刻的序号水位 / Sequence watermark at the last acknowledge
    uFirstSeq     : UDINT;                  // 扫描中的首出候选序号 / First-out candidate sequence during the scan
    uTopSeq       : UDINT;                  // 扫描中的最高优先级候选序号 / Top-priority candidate sequence during the scan
    bLatchValid   : BOOL;                   // 首出锁存有效 / First-out latch valid
    fbTrigAck     : R_TRIG;                 // 确认上升沿检测实例 / Acknowledge rising edge detector instance
    nIdx          : INT;                    // 扫描索引，值域 0..15 / Scan index, range 0..15
    nBestPrio     : USINT;                  // 扫描中的最优优先级 / Best priority during the scan
    uBestSeq      : UDINT;                  // 扫描中的最优序号（保留诊断口径）/ Best sequence during the scan
END_VAR
VAR CONSTANT
    DL_ALM_CH_COUNT  : INT   := 16;             // 通道数 [个]，与数组维度一致 / Channel count [count], must match the arrays
    DL_ALM_PRIO_STOP : USINT := 1;              // 停机级 / Stop level
    DL_ALM_PRIO_WARN : USINT := 2;              // 警告级 / Warning level
    DL_ALM_PRIO_INFO : USINT := 3;              // 提示级 / Info level
    DL_ALM_PRIO_MAX  : USINT := 3;              // 合法优先级上限 / Max valid priority
    DL_ALM_IDX_NONE  : INT   := -1;             // 无效通道索引哨兵 / Sentinel for no channel
    DL_ALM_SEQ_MAX   : UDINT := 16#FFFF_FFFE;   // 序号饱和上限，不回绕 / Sequence saturation limit, no wrap-around
END_VAR

(*------------------------------------------------------------------------------
 * 段 1｜无条件刷新区（红线 R7）：确认沿实例位于主体最前部，严禁进入 IF / CASE
 *      Unconditional refresh zone: the acknowledge edge instance runs at the very top
 *-----------------------------------------------------------------------------*)
fbTrigAck(CLK := bAck);

(*------------------------------------------------------------------------------
 * 段 2｜故障码本周期清零
 *      Error code is cleared every scan
 *-----------------------------------------------------------------------------*)
uErrorId := 16#0000_0000;

(*------------------------------------------------------------------------------
 * 段 3｜使能失效（决策 P6）：输出与序号表全部清零，重新使能视同冷启动
 *      Disabled: outputs and the sequence table are cleared, re-enable is a cold start
 *-----------------------------------------------------------------------------*)
IF NOT bEnable THEN

    uAlarmWord   := 16#0000;
    uActiveCount := USINT#0;
    bAnyActive   := FALSE;
    bShutdown    := FALSE;
    nFirstOutIdx := DL_ALM_IDX_NONE;
    bFirstOutAck := FALSE;
    nTopPrioIdx  := DL_ALM_IDX_NONE;
    bLatchValid  := FALSE;
    uSeqNext     := UDINT#0;
    uAckSeq      := UDINT#0;

    FOR nIdx := 0 TO (DL_ALM_CH_COUNT - 1) DO
        IF (nIdx >= 0) AND (nIdx < DL_ALM_CH_COUNT) THEN
            auSeqNo[nIdx]   := UDINT#0;
            auPrioEff[nIdx] := USINT#0;
            abPackSrc[nIdx] := FALSE;
        END_IF
    END_FOR;

ELSE

    (*--------------------------------------------------------------------------
     * 段 4｜确认水位推进（边界 B5）：确认沿只推水位，绝不动激活态
     *      Acknowledge: advance the watermark only, the active states are untouched
     *-------------------------------------------------------------------------*)
    IF fbTrigAck.Q THEN
        uAckSeq := uSeqNext;
    END_IF

    (*--------------------------------------------------------------------------
     * 段 5｜优先级钳位与激活取号（边界 B2/B3/B6/B9）：单次全通道扫描完成
     *      Priority clamp and activation numbering in one full-channel scan
     *      激活沿取号：通道由未激活变激活时取当前序号并递增发生器
     *      Activation numbering: a channel takes a number when it starts alarming
     *      通道消失即清号，使其下次激活能重新排队参与首出竞争
     *      The number is cleared on deactivation so a re-activation queues again
     *-------------------------------------------------------------------------*)
    FOR nIdx := 0 TO (DL_ALM_CH_COUNT - 1) DO

        IF (nIdx >= 0) AND (nIdx < DL_ALM_CH_COUNT) THEN

            IF auPriority[nIdx] > DL_ALM_PRIO_MAX THEN
                auPrioEff[nIdx] := DL_ALM_PRIO_MAX;
                uErrorId        := 16#0001_0001;
            ELSE
                auPrioEff[nIdx] := auPriority[nIdx];
            END_IF

            IF abAlarmActive[nIdx] THEN
                IF auSeqNo[nIdx] = UDINT#0 THEN
                    IF uSeqNext < DL_ALM_SEQ_MAX THEN
                        uSeqNext        := uSeqNext + UDINT#1;
                        auSeqNo[nIdx]   := uSeqNext;
                    ELSE
                        (* 序号饱和停增：回绕会破坏先到先得次序（边界 B6） *)
                        (* Saturation instead of wrap-around keeps the arrival order intact *)
                        auSeqNo[nIdx] := DL_ALM_SEQ_MAX;
                        uErrorId      := 16#0001_0007;
                    END_IF
                END_IF
            ELSE
                auSeqNo[nIdx] := UDINT#0;
            END_IF

        END_IF

    END_FOR;

    (*--------------------------------------------------------------------------
     * 段 6｜仲裁扫描（边界 B4）：首出取最小序号，最高优先级取最小优先级
     *      Arbitration: first-out is the smallest sequence, top priority the smallest level
     *      同级之间再比序号，实现"同级先到先得"，扫描为有限 FOR，无 WHILE
     *      Ties are broken by the sequence number, the scan is a bounded FOR loop
     *-------------------------------------------------------------------------*)
    nFirstOutIdx := DL_ALM_IDX_NONE;
    nTopPrioIdx  := DL_ALM_IDX_NONE;
    nBestPrio    := DL_ALM_PRIO_MAX;
    uFirstSeq    := UDINT#0;
    uTopSeq      := UDINT#0;
    uBestSeq     := UDINT#0;
    uActiveCount := USINT#0;
    bShutdown    := FALSE;

    FOR nIdx := 0 TO (DL_ALM_CH_COUNT - 1) DO

        IF (nIdx >= 0) AND (nIdx < DL_ALM_CH_COUNT) THEN

            (* 禁用通道（优先级 0）不参与计数与仲裁 *)
            (* Disabled channels take no part in counting or arbitration *)
            IF abAlarmActive[nIdx] AND (auPrioEff[nIdx] > USINT#0) THEN

                uActiveCount := uActiveCount + USINT#1;

                IF auPrioEff[nIdx] = DL_ALM_PRIO_STOP THEN
                    bShutdown := TRUE;
                END_IF

                (*--------------------------------------------------------------
                 * 段 6a｜首出候选：只接受晚于确认水位的序号（已确认的不再补位）
                 *      First-out candidate: only sequences newer than the watermark count
                 *-------------------------------------------------------------*)
                IF auSeqNo[nIdx] > uAckSeq THEN
                    IF (nFirstOutIdx = DL_ALM_IDX_NONE) OR (auSeqNo[nIdx] < uFirstSeq) THEN
                        nFirstOutIdx := nIdx;
                        uFirstSeq    := auSeqNo[nIdx];
                    END_IF
                END_IF

                (*--------------------------------------------------------------
                 * 段 6b｜最高优先级候选：优先级数值更小者胜，同级比序号
                 *      Top-priority candidate: the smaller level wins, ties by sequence
                 *-------------------------------------------------------------*)
                IF (nTopPrioIdx = DL_ALM_IDX_NONE) OR (auPrioEff[nIdx] < nBestPrio) THEN
                    nTopPrioIdx := nIdx;
                    nBestPrio   := auPrioEff[nIdx];
                    uTopSeq     := auSeqNo[nIdx];
                    uBestSeq    := auSeqNo[nIdx];
                ELSIF (auPrioEff[nIdx] = nBestPrio) AND (auSeqNo[nIdx] < uTopSeq) THEN
                    nTopPrioIdx := nIdx;
                    uTopSeq     := auSeqNo[nIdx];
                END_IF

            END_IF

        END_IF

    END_FOR;

    (*--------------------------------------------------------------------------
     * 段 7｜报警字打包（边界 B7）：先构造打包源，再调用位打包构件
     *      Bitmap packing: build the source array first, then call the packing function
     *      禁用通道对应位强制 0：报警字是给上位机的最终事实，
     *      混入"禁用但确实跳了"的位会让上位机与 PLC 状态产生错觉（决策 P5）
     *      Disabled bits are forced to zero so the bitmap never contradicts the arbitration
     *-------------------------------------------------------------------------*)
    FOR nIdx := 0 TO (DL_ALM_CH_COUNT - 1) DO
        IF (nIdx >= 0) AND (nIdx < DL_ALM_CH_COUNT) THEN
            abPackSrc[nIdx] := abAlarmActive[nIdx] AND (auPrioEff[nIdx] > USINT#0);
        END_IF
    END_FOR;

    uAlarmWord := FC_DL_PackBitsToWord(abBits := abPackSrc);

    (*--------------------------------------------------------------------------
     * 段 8｜输出汇总（边界 B5）：三态正交——激活、已确认、首出锁存各管一路
     *      Output summary: active, acknowledged and first-out latched stay orthogonal
     *-------------------------------------------------------------------------*)
    bLatchValid  := (nFirstOutIdx <> DL_ALM_IDX_NONE);
    bAnyActive   := (uActiveCount > USINT#0);
    bFirstOutAck := (NOT bLatchValid) AND (uAckSeq > UDINT#0);

END_IF
END_FUNCTION_BLOCK
